REGION Network 31: Level Conveyors Tower 2 - SYSTEM 3
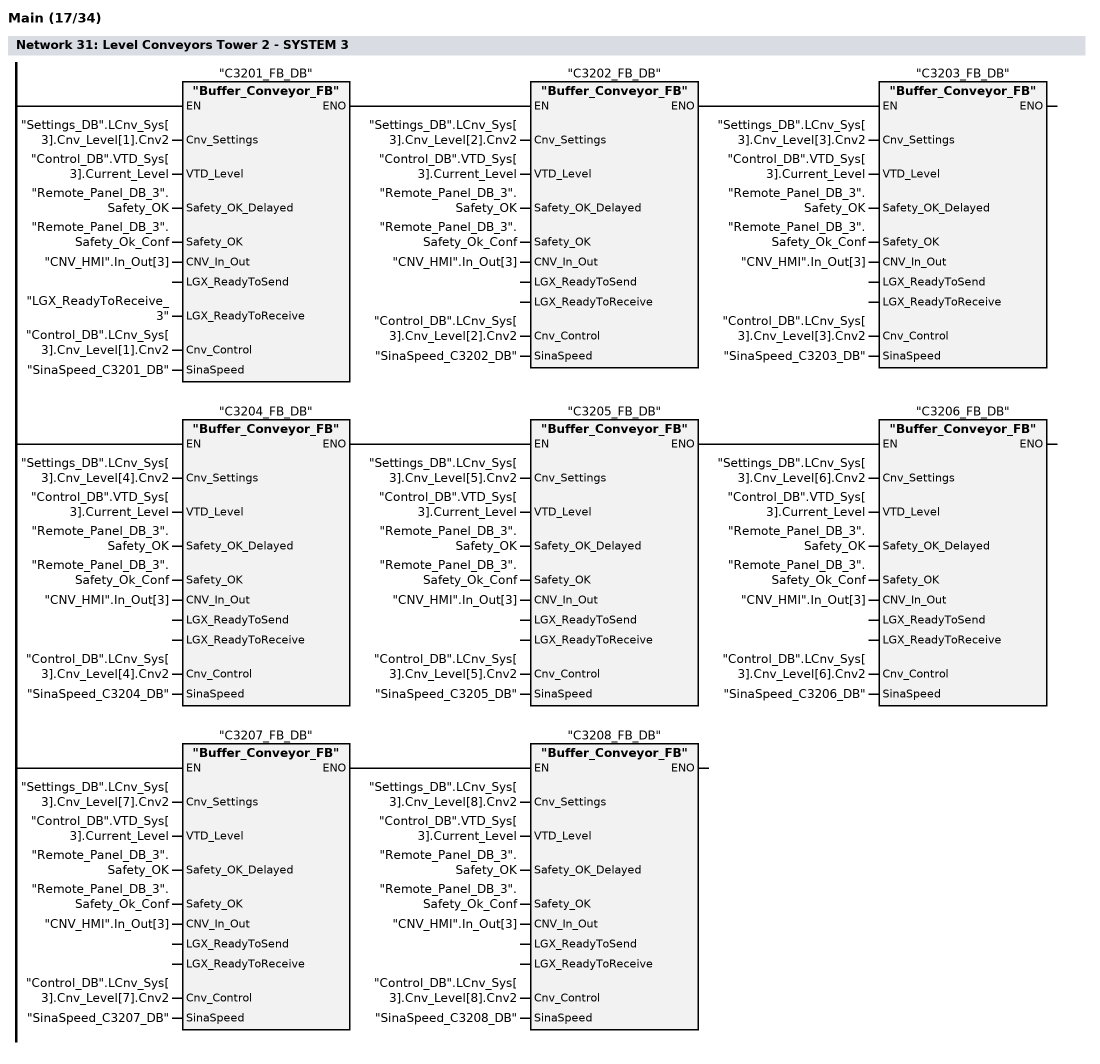
   RUNG wire#powerrail
      "C3201_FB_DB"(Cnv_Settings := "Settings_DB".LCnv_Sys[3].Cnv_Level[1].Cnv2, VTD_Level := "Control_DB".VTD_Sys[3].Current_Level, Safety_OK_Delayed := "Remote_Panel_DB_3".Safety_OK, Safety_OK := "Remote_Panel_DB_3".Safety_Ok_Conf, CNV_In_Out := "CNV_HMI".In_Out[3], LGX_ReadyToSend :=, LGX_ReadyToReceive := "LGX_ReadyToReceive_3", Cnv_Control := "Control_DB".LCnv_Sys[3].Cnv_Level[1].Cnv2, SinaSpeed := "SinaSpeed_C3201_DB")
      "C3202_FB_DB"(Cnv_Settings := "Settings_DB".LCnv_Sys[3].Cnv_Level[2].Cnv2, VTD_Level := "Control_DB".VTD_Sys[3].Current_Level, Safety_OK_Delayed := "Remote_Panel_DB_3".Safety_OK, Safety_OK := "Remote_Panel_DB_3".Safety_Ok_Conf, CNV_In_Out := "CNV_HMI".In_Out[3], LGX_ReadyToSend :=, LGX_ReadyToReceive :=, Cnv_Control := "Control_DB".LCnv_Sys[3].Cnv_Level[2].Cnv2, SinaSpeed := "SinaSpeed_C3202_DB")
      "C3203_FB_DB"(Cnv_Settings := "Settings_DB".LCnv_Sys[3].Cnv_Level[3].Cnv2, VTD_Level := "Control_DB".VTD_Sys[3].Current_Level, Safety_OK_Delayed := "Remote_Panel_DB_3".Safety_OK, Safety_OK := "Remote_Panel_DB_3".Safety_Ok_Conf, CNV_In_Out := "CNV_HMI".In_Out[3], LGX_ReadyToSend :=, LGX_ReadyToReceive :=, Cnv_Control := "Control_DB".LCnv_Sys[3].Cnv_Level[3].Cnv2, SinaSpeed := "SinaSpeed_C3203_DB")
   END_RUNG
   RUNG wire#powerrail
      "C3204_FB_DB"(Cnv_Settings := "Settings_DB".LCnv_Sys[3].Cnv_Level[4].Cnv2, VTD_Level := "Control_DB".VTD_Sys[3].Current_Level, Safety_OK_Delayed := "Remote_Panel_DB_3".Safety_OK, Safety_OK := "Remote_Panel_DB_3".Safety_Ok_Conf, CNV_In_Out := "CNV_HMI".In_Out[3], LGX_ReadyToSend :=, LGX_ReadyToReceive :=, Cnv_Control := "Control_DB".LCnv_Sys[3].Cnv_Level[4].Cnv2, SinaSpeed := "SinaSpeed_C3204_DB")
      "C3205_FB_DB"(Cnv_Settings := "Settings_DB".LCnv_Sys[3].Cnv_Level[5].Cnv2, VTD_Level := "Control_DB".VTD_Sys[3].Current_Level, Safety_OK_Delayed := "Remote_Panel_DB_3".Safety_OK, Safety_OK := "Remote_Panel_DB_3".Safety_Ok_Conf, CNV_In_Out := "CNV_HMI".In_Out[3], LGX_ReadyToSend :=, LGX_ReadyToReceive :=, Cnv_Control := "Control_DB".LCnv_Sys[3].Cnv_Level[5].Cnv2, SinaSpeed := "SinaSpeed_C3205_DB")
      "C3206_FB_DB"(Cnv_Settings := "Settings_DB".LCnv_Sys[3].Cnv_Level[6].Cnv2, VTD_Level := "Control_DB".VTD_Sys[3].Current_Level, Safety_OK_Delayed := "Remote_Panel_DB_3".Safety_OK, Safety_OK := "Remote_Panel_DB_3".Safety_Ok_Conf, CNV_In_Out := "CNV_HMI".In_Out[3], LGX_ReadyToSend :=, LGX_ReadyToReceive :=, Cnv_Control := "Control_DB".LCnv_Sys[3].Cnv_Level[6].Cnv2, SinaSpeed := "SinaSpeed_C3206_DB")
   END_RUNG
   RUNG wire#powerrail
      "C3207_FB_DB"(Cnv_Settings := "Settings_DB".LCnv_Sys[3].Cnv_Level[7].Cnv2, VTD_Level := "Control_DB".VTD_Sys[3].Current_Level, Safety_OK_Delayed := "Remote_Panel_DB_3".Safety_OK, Safety_OK := "Remote_Panel_DB_3".Safety_Ok_Conf, CNV_In_Out := "CNV_HMI".In_Out[3], LGX_ReadyToSend :=, LGX_ReadyToReceive :=, Cnv_Control := "Control_DB".LCnv_Sys[3].Cnv_Level[7].Cnv2, SinaSpeed := "SinaSpeed_C3207_DB")
      "C3208_FB_DB"(Cnv_Settings := "Settings_DB".LCnv_Sys[3].Cnv_Level[8].Cnv2, VTD_Level := "Control_DB".VTD_Sys[3].Current_Level, Safety_OK_Delayed := "Remote_Panel_DB_3".Safety_OK, Safety_OK := "Remote_Panel_DB_3".Safety_Ok_Conf, CNV_In_Out := "CNV_HMI".In_Out[3], LGX_ReadyToSend :=, LGX_ReadyToReceive :=, Cnv_Control := "Control_DB".LCnv_Sys[3].Cnv_Level[8].Cnv2, SinaSpeed := "SinaSpeed_C3208_DB")
   END_RUNG
   // the same network as SCL:
   "C3201_FB_DB"(Cnv_Settings := "Settings_DB".LCnv_Sys[3].Cnv_Level[1].Cnv2,   // "Buffer_Conveyor_FB"
                 VTD_Level := "Control_DB".VTD_Sys[3].Current_Level,
                 Safety_OK_Delayed := "Remote_Panel_DB_3".Safety_OK,
                 Safety_OK := "Remote_Panel_DB_3".Safety_Ok_Conf,
                 CNV_In_Out := "CNV_HMI".In_Out[3],
                 LGX_ReadyToReceive := "LGX_ReadyToReceive_3",
                 Cnv_Control := "Control_DB".LCnv_Sys[3].Cnv_Level[1].Cnv2,
                 SinaSpeed := "SinaSpeed_C3201_DB",
                 ENO => #_w1);
   "C3202_FB_DB"(EN := #_w1,   // "Buffer_Conveyor_FB"
                 Cnv_Settings := "Settings_DB".LCnv_Sys[3].Cnv_Level[2].Cnv2,
                 VTD_Level := "Control_DB".VTD_Sys[3].Current_Level,
                 Safety_OK_Delayed := "Remote_Panel_DB_3".Safety_OK,
                 Safety_OK := "Remote_Panel_DB_3".Safety_Ok_Conf,
                 CNV_In_Out := "CNV_HMI".In_Out[3],
                 Cnv_Control := "Control_DB".LCnv_Sys[3].Cnv_Level[2].Cnv2,
                 SinaSpeed := "SinaSpeed_C3202_DB",
                 ENO => #_w2);
   IF #_w2 THEN
       "C3203_FB_DB"(Cnv_Settings := "Settings_DB".LCnv_Sys[3].Cnv_Level[3].Cnv2,   // "Buffer_Conveyor_FB"
                     VTD_Level := "Control_DB".VTD_Sys[3].Current_Level,
                     Safety_OK_Delayed := "Remote_Panel_DB_3".Safety_OK,
                     Safety_OK := "Remote_Panel_DB_3".Safety_Ok_Conf,
                     CNV_In_Out := "CNV_HMI".In_Out[3],
                     Cnv_Control := "Control_DB".LCnv_Sys[3].Cnv_Level[3].Cnv2,
                     SinaSpeed := "SinaSpeed_C3203_DB");
   END_IF;
   "C3204_FB_DB"(Cnv_Settings := "Settings_DB".LCnv_Sys[3].Cnv_Level[4].Cnv2,   // "Buffer_Conveyor_FB"
                 VTD_Level := "Control_DB".VTD_Sys[3].Current_Level,
                 Safety_OK_Delayed := "Remote_Panel_DB_3".Safety_OK,
                 Safety_OK := "Remote_Panel_DB_3".Safety_Ok_Conf,
                 CNV_In_Out := "CNV_HMI".In_Out[3],
                 Cnv_Control := "Control_DB".LCnv_Sys[3].Cnv_Level[4].Cnv2,
                 SinaSpeed := "SinaSpeed_C3204_DB",
                 ENO => #_w3);
   "C3205_FB_DB"(EN := #_w3,   // "Buffer_Conveyor_FB"
                 Cnv_Settings := "Settings_DB".LCnv_Sys[3].Cnv_Level[5].Cnv2,
                 VTD_Level := "Control_DB".VTD_Sys[3].Current_Level,
                 Safety_OK_Delayed := "Remote_Panel_DB_3".Safety_OK,
                 Safety_OK := "Remote_Panel_DB_3".Safety_Ok_Conf,
                 CNV_In_Out := "CNV_HMI".In_Out[3],
                 Cnv_Control := "Control_DB".LCnv_Sys[3].Cnv_Level[5].Cnv2,
                 SinaSpeed := "SinaSpeed_C3205_DB",
                 ENO => #_w4);
   IF #_w4 THEN
       "C3206_FB_DB"(Cnv_Settings := "Settings_DB".LCnv_Sys[3].Cnv_Level[6].Cnv2,   // "Buffer_Conveyor_FB"
                     VTD_Level := "Control_DB".VTD_Sys[3].Current_Level,
                     Safety_OK_Delayed := "Remote_Panel_DB_3".Safety_OK,
                     Safety_OK := "Remote_Panel_DB_3".Safety_Ok_Conf,
                     CNV_In_Out := "CNV_HMI".In_Out[3],
                     Cnv_Control := "Control_DB".LCnv_Sys[3].Cnv_Level[6].Cnv2,
                     SinaSpeed := "SinaSpeed_C3206_DB");
   END_IF;
   "C3207_FB_DB"(Cnv_Settings := "Settings_DB".LCnv_Sys[3].Cnv_Level[7].Cnv2,   // "Buffer_Conveyor_FB"
                 VTD_Level := "Control_DB".VTD_Sys[3].Current_Level,
                 Safety_OK_Delayed := "Remote_Panel_DB_3".Safety_OK,
                 Safety_OK := "Remote_Panel_DB_3".Safety_Ok_Conf,
                 CNV_In_Out := "CNV_HMI".In_Out[3],
                 Cnv_Control := "Control_DB".LCnv_Sys[3].Cnv_Level[7].Cnv2,
                 SinaSpeed := "SinaSpeed_C3207_DB",
                 ENO => #_w5);
   IF #_w5 THEN
       "C3208_FB_DB"(Cnv_Settings := "Settings_DB".LCnv_Sys[3].Cnv_Level[8].Cnv2,   // "Buffer_Conveyor_FB"
                     VTD_Level := "Control_DB".VTD_Sys[3].Current_Level,
                     Safety_OK_Delayed := "Remote_Panel_DB_3".Safety_OK,
                     Safety_OK := "Remote_Panel_DB_3".Safety_Ok_Conf,
                     CNV_In_Out := "CNV_HMI".In_Out[3],
                     Cnv_Control := "Control_DB".LCnv_Sys[3].Cnv_Level[8].Cnv2,
                     SinaSpeed := "SinaSpeed_C3208_DB");
   END_IF;
END_REGION

REGION Network 32: SAFETY STOPPERS Tower 1 - SYSTEM 3
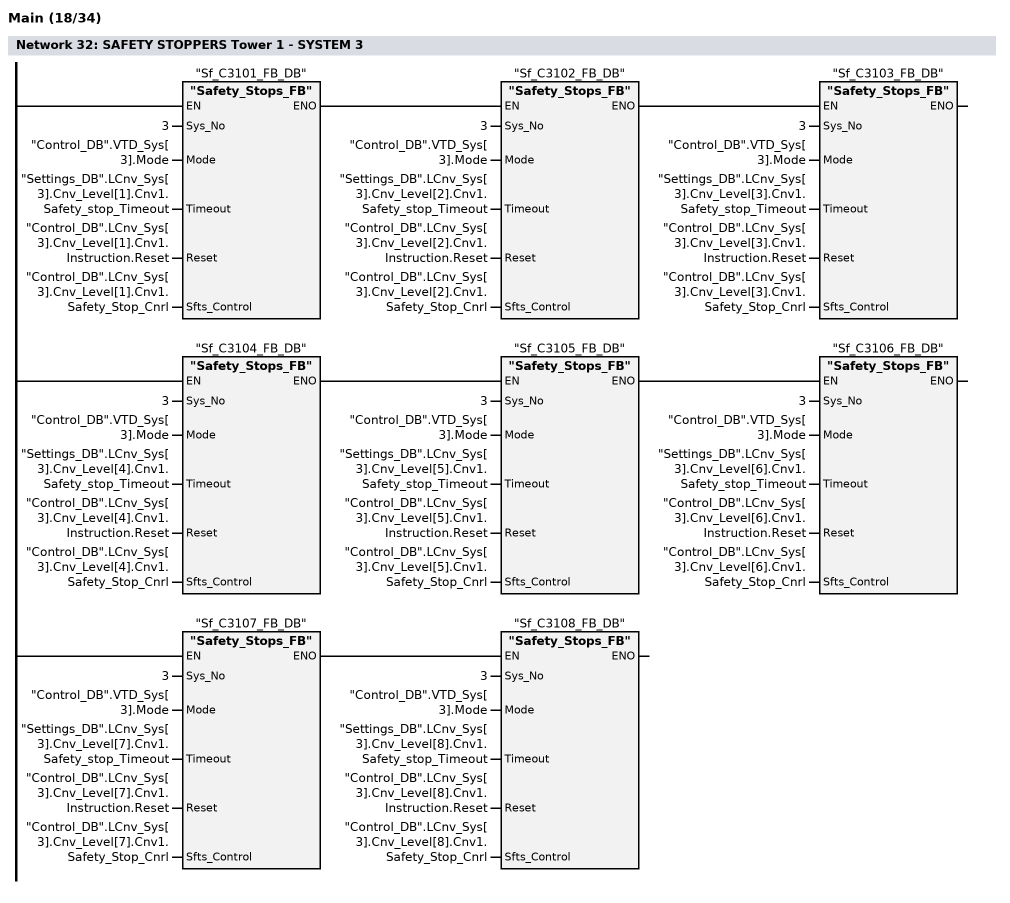
   RUNG wire#powerrail
      "Sf_C3101_FB_DB"(Sys_No := 3, Mode := "Control_DB".VTD_Sys[3].Mode, Timeout := "Settings_DB".LCnv_Sys[3].Cnv_Level[1].Cnv1.Safety_stop_Timeout, Reset := "Control_DB".LCnv_Sys[3].Cnv_Level[1].Cnv1.Instruction.Reset, Sfts_Control := "Control_DB".LCnv_Sys[3].Cnv_Level[1].Cnv1.Safety_Stop_Cnrl)
      "Sf_C3102_FB_DB"(Sys_No := 3, Mode := "Control_DB".VTD_Sys[3].Mode, Timeout := "Settings_DB".LCnv_Sys[3].Cnv_Level[2].Cnv1.Safety_stop_Timeout, Reset := "Control_DB".LCnv_Sys[3].Cnv_Level[2].Cnv1.Instruction.Reset, Sfts_Control := "Control_DB".LCnv_Sys[3].Cnv_Level[2].Cnv1.Safety_Stop_Cnrl)
      "Sf_C3103_FB_DB"(Sys_No := 3, Mode := "Control_DB".VTD_Sys[3].Mode, Timeout := "Settings_DB".LCnv_Sys[3].Cnv_Level[3].Cnv1.Safety_stop_Timeout, Reset := "Control_DB".LCnv_Sys[3].Cnv_Level[3].Cnv1.Instruction.Reset, Sfts_Control := "Control_DB".LCnv_Sys[3].Cnv_Level[3].Cnv1.Safety_Stop_Cnrl)
   END_RUNG
   RUNG wire#powerrail
      "Sf_C3104_FB_DB"(Sys_No := 3, Mode := "Control_DB".VTD_Sys[3].Mode, Timeout := "Settings_DB".LCnv_Sys[3].Cnv_Level[4].Cnv1.Safety_stop_Timeout, Reset := "Control_DB".LCnv_Sys[3].Cnv_Level[4].Cnv1.Instruction.Reset, Sfts_Control := "Control_DB".LCnv_Sys[3].Cnv_Level[4].Cnv1.Safety_Stop_Cnrl)
      "Sf_C3105_FB_DB"(Sys_No := 3, Mode := "Control_DB".VTD_Sys[3].Mode, Timeout := "Settings_DB".LCnv_Sys[3].Cnv_Level[5].Cnv1.Safety_stop_Timeout, Reset := "Control_DB".LCnv_Sys[3].Cnv_Level[5].Cnv1.Instruction.Reset, Sfts_Control := "Control_DB".LCnv_Sys[3].Cnv_Level[5].Cnv1.Safety_Stop_Cnrl)
      "Sf_C3106_FB_DB"(Sys_No := 3, Mode := "Control_DB".VTD_Sys[3].Mode, Timeout := "Settings_DB".LCnv_Sys[3].Cnv_Level[6].Cnv1.Safety_stop_Timeout, Reset := "Control_DB".LCnv_Sys[3].Cnv_Level[6].Cnv1.Instruction.Reset, Sfts_Control := "Control_DB".LCnv_Sys[3].Cnv_Level[6].Cnv1.Safety_Stop_Cnrl)
   END_RUNG
   RUNG wire#powerrail
      "Sf_C3107_FB_DB"(Sys_No := 3, Mode := "Control_DB".VTD_Sys[3].Mode, Timeout := "Settings_DB".LCnv_Sys[3].Cnv_Level[7].Cnv1.Safety_stop_Timeout, Reset := "Control_DB".LCnv_Sys[3].Cnv_Level[7].Cnv1.Instruction.Reset, Sfts_Control := "Control_DB".LCnv_Sys[3].Cnv_Level[7].Cnv1.Safety_Stop_Cnrl)
      "Sf_C3108_FB_DB"(Sys_No := 3, Mode := "Control_DB".VTD_Sys[3].Mode, Timeout := "Settings_DB".LCnv_Sys[3].Cnv_Level[8].Cnv1.Safety_stop_Timeout, Reset := "Control_DB".LCnv_Sys[3].Cnv_Level[8].Cnv1.Instruction.Reset, Sfts_Control := "Control_DB".LCnv_Sys[3].Cnv_Level[8].Cnv1.Safety_Stop_Cnrl)
   END_RUNG
   // the same network as SCL:
   "Sf_C3101_FB_DB"(Sys_No := 3,   // "Safety_Stops_FB"
                    Mode := "Control_DB".VTD_Sys[3].Mode,
                    Timeout := "Settings_DB".LCnv_Sys[3].Cnv_Level[1].Cnv1.Safety_stop_Timeout,
                    Reset := "Control_DB".LCnv_Sys[3].Cnv_Level[1].Cnv1.Instruction.Reset,
                    Sfts_Control := "Control_DB".LCnv_Sys[3].Cnv_Level[1].Cnv1.Safety_Stop_Cnrl,
                    ENO => #_w1);
   "Sf_C3102_FB_DB"(EN := #_w1,   // "Safety_Stops_FB"
                    Sys_No := 3,
                    Mode := "Control_DB".VTD_Sys[3].Mode,
                    Timeout := "Settings_DB".LCnv_Sys[3].Cnv_Level[2].Cnv1.Safety_stop_Timeout,
                    Reset := "Control_DB".LCnv_Sys[3].Cnv_Level[2].Cnv1.Instruction.Reset,
                    Sfts_Control := "Control_DB".LCnv_Sys[3].Cnv_Level[2].Cnv1.Safety_Stop_Cnrl,
                    ENO => #_w2);
   IF #_w2 THEN
       "Sf_C3103_FB_DB"(Sys_No := 3,   // "Safety_Stops_FB"
                        Mode := "Control_DB".VTD_Sys[3].Mode,
                        Timeout := "Settings_DB".LCnv_Sys[3].Cnv_Level[3].Cnv1.Safety_stop_Timeout,
                        Reset := "Control_DB".LCnv_Sys[3].Cnv_Level[3].Cnv1.Instruction.Reset,
                        Sfts_Control := "Control_DB".LCnv_Sys[3].Cnv_Level[3].Cnv1.Safety_Stop_Cnrl);
   END_IF;
   "Sf_C3104_FB_DB"(Sys_No := 3,   // "Safety_Stops_FB"
                    Mode := "Control_DB".VTD_Sys[3].Mode,
                    Timeout := "Settings_DB".LCnv_Sys[3].Cnv_Level[4].Cnv1.Safety_stop_Timeout,
                    Reset := "Control_DB".LCnv_Sys[3].Cnv_Level[4].Cnv1.Instruction.Reset,
                    Sfts_Control := "Control_DB".LCnv_Sys[3].Cnv_Level[4].Cnv1.Safety_Stop_Cnrl,
                    ENO => #_w3);
   "Sf_C3105_FB_DB"(EN := #_w3,   // "Safety_Stops_FB"
                    Sys_No := 3,
                    Mode := "Control_DB".VTD_Sys[3].Mode,
                    Timeout := "Settings_DB".LCnv_Sys[3].Cnv_Level[5].Cnv1.Safety_stop_Timeout,
                    Reset := "Control_DB".LCnv_Sys[3].Cnv_Level[5].Cnv1.Instruction.Reset,
                    Sfts_Control := "Control_DB".LCnv_Sys[3].Cnv_Level[5].Cnv1.Safety_Stop_Cnrl,
                    ENO => #_w4);
   IF #_w4 THEN
       "Sf_C3106_FB_DB"(Sys_No := 3,   // "Safety_Stops_FB"
                        Mode := "Control_DB".VTD_Sys[3].Mode,
                        Timeout := "Settings_DB".LCnv_Sys[3].Cnv_Level[6].Cnv1.Safety_stop_Timeout,
                        Reset := "Control_DB".LCnv_Sys[3].Cnv_Level[6].Cnv1.Instruction.Reset,
                        Sfts_Control := "Control_DB".LCnv_Sys[3].Cnv_Level[6].Cnv1.Safety_Stop_Cnrl);
   END_IF;
   "Sf_C3107_FB_DB"(Sys_No := 3,   // "Safety_Stops_FB"
                    Mode := "Control_DB".VTD_Sys[3].Mode,
                    Timeout := "Settings_DB".LCnv_Sys[3].Cnv_Level[7].Cnv1.Safety_stop_Timeout,
                    Reset := "Control_DB".LCnv_Sys[3].Cnv_Level[7].Cnv1.Instruction.Reset,
                    Sfts_Control := "Control_DB".LCnv_Sys[3].Cnv_Level[7].Cnv1.Safety_Stop_Cnrl,
                    ENO => #_w5);
   IF #_w5 THEN
       "Sf_C3108_FB_DB"(Sys_No := 3,   // "Safety_Stops_FB"
                        Mode := "Control_DB".VTD_Sys[3].Mode,
                        Timeout := "Settings_DB".LCnv_Sys[3].Cnv_Level[8].Cnv1.Safety_stop_Timeout,
                        Reset := "Control_DB".LCnv_Sys[3].Cnv_Level[8].Cnv1.Instruction.Reset,
                        Sfts_Control := "Control_DB".LCnv_Sys[3].Cnv_Level[8].Cnv1.Safety_Stop_Cnrl);
   END_IF;
END_REGION

REGION Network 33: SAFETY STOPPERS Tower 2 - SYSTEM 3
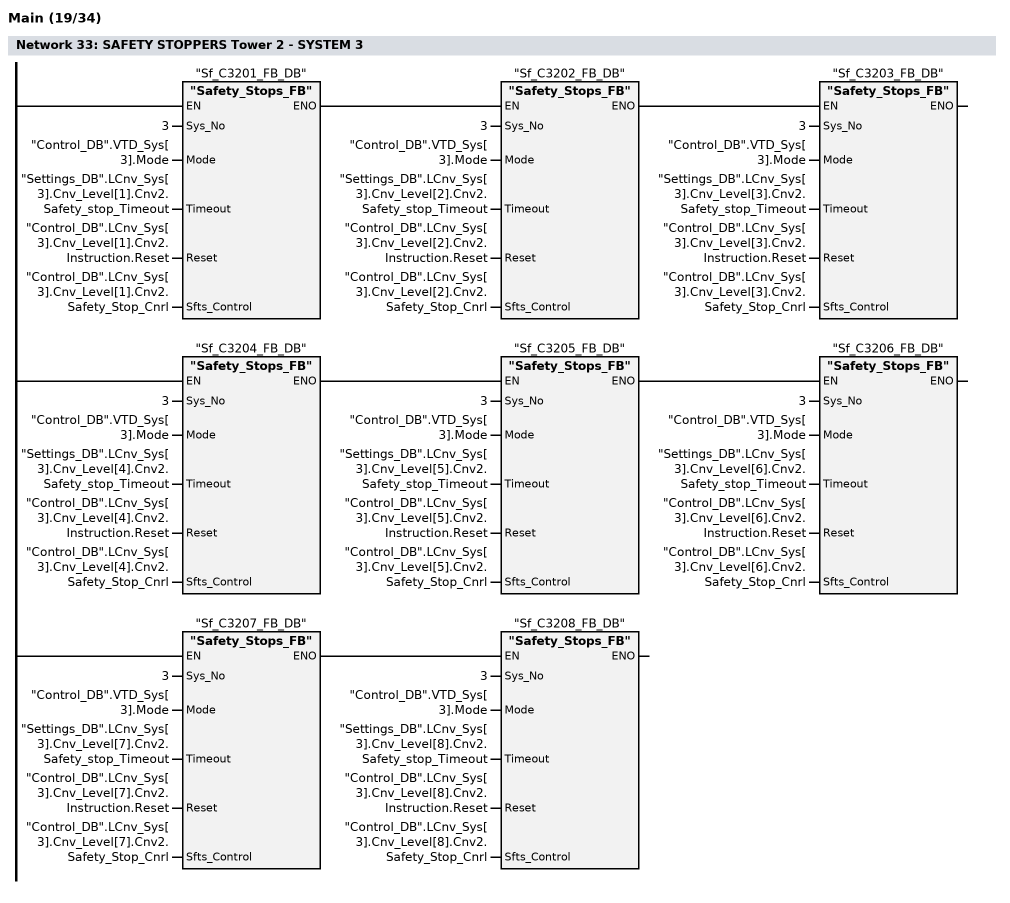
   RUNG wire#powerrail
      "Sf_C3201_FB_DB"(Sys_No := 3, Mode := "Control_DB".VTD_Sys[3].Mode, Timeout := "Settings_DB".LCnv_Sys[3].Cnv_Level[1].Cnv2.Safety_stop_Timeout, Reset := "Control_DB".LCnv_Sys[3].Cnv_Level[1].Cnv2.Instruction.Reset, Sfts_Control := "Control_DB".LCnv_Sys[3].Cnv_Level[1].Cnv2.Safety_Stop_Cnrl)
      "Sf_C3202_FB_DB"(Sys_No := 3, Mode := "Control_DB".VTD_Sys[3].Mode, Timeout := "Settings_DB".LCnv_Sys[3].Cnv_Level[2].Cnv2.Safety_stop_Timeout, Reset := "Control_DB".LCnv_Sys[3].Cnv_Level[2].Cnv2.Instruction.Reset, Sfts_Control := "Control_DB".LCnv_Sys[3].Cnv_Level[2].Cnv2.Safety_Stop_Cnrl)
      "Sf_C3203_FB_DB"(Sys_No := 3, Mode := "Control_DB".VTD_Sys[3].Mode, Timeout := "Settings_DB".LCnv_Sys[3].Cnv_Level[3].Cnv2.Safety_stop_Timeout, Reset := "Control_DB".LCnv_Sys[3].Cnv_Level[3].Cnv2.Instruction.Reset, Sfts_Control := "Control_DB".LCnv_Sys[3].Cnv_Level[3].Cnv2.Safety_Stop_Cnrl)
   END_RUNG
   RUNG wire#powerrail
      "Sf_C3204_FB_DB"(Sys_No := 3, Mode := "Control_DB".VTD_Sys[3].Mode, Timeout := "Settings_DB".LCnv_Sys[3].Cnv_Level[4].Cnv2.Safety_stop_Timeout, Reset := "Control_DB".LCnv_Sys[3].Cnv_Level[4].Cnv2.Instruction.Reset, Sfts_Control := "Control_DB".LCnv_Sys[3].Cnv_Level[4].Cnv2.Safety_Stop_Cnrl)
      "Sf_C3205_FB_DB"(Sys_No := 3, Mode := "Control_DB".VTD_Sys[3].Mode, Timeout := "Settings_DB".LCnv_Sys[3].Cnv_Level[5].Cnv2.Safety_stop_Timeout, Reset := "Control_DB".LCnv_Sys[3].Cnv_Level[5].Cnv2.Instruction.Reset, Sfts_Control := "Control_DB".LCnv_Sys[3].Cnv_Level[5].Cnv2.Safety_Stop_Cnrl)
      "Sf_C3206_FB_DB"(Sys_No := 3, Mode := "Control_DB".VTD_Sys[3].Mode, Timeout := "Settings_DB".LCnv_Sys[3].Cnv_Level[6].Cnv2.Safety_stop_Timeout, Reset := "Control_DB".LCnv_Sys[3].Cnv_Level[6].Cnv2.Instruction.Reset, Sfts_Control := "Control_DB".LCnv_Sys[3].Cnv_Level[6].Cnv2.Safety_Stop_Cnrl)
   END_RUNG
   RUNG wire#powerrail
      "Sf_C3207_FB_DB"(Sys_No := 3, Mode := "Control_DB".VTD_Sys[3].Mode, Timeout := "Settings_DB".LCnv_Sys[3].Cnv_Level[7].Cnv2.Safety_stop_Timeout, Reset := "Control_DB".LCnv_Sys[3].Cnv_Level[7].Cnv2.Instruction.Reset, Sfts_Control := "Control_DB".LCnv_Sys[3].Cnv_Level[7].Cnv2.Safety_Stop_Cnrl)
      "Sf_C3208_FB_DB"(Sys_No := 3, Mode := "Control_DB".VTD_Sys[3].Mode, Timeout := "Settings_DB".LCnv_Sys[3].Cnv_Level[8].Cnv2.Safety_stop_Timeout, Reset := "Control_DB".LCnv_Sys[3].Cnv_Level[8].Cnv2.Instruction.Reset, Sfts_Control := "Control_DB".LCnv_Sys[3].Cnv_Level[8].Cnv2.Safety_Stop_Cnrl)
   END_RUNG
   // the same network as SCL:
   "Sf_C3201_FB_DB"(Sys_No := 3,   // "Safety_Stops_FB"
                    Mode := "Control_DB".VTD_Sys[3].Mode,
                    Timeout := "Settings_DB".LCnv_Sys[3].Cnv_Level[1].Cnv2.Safety_stop_Timeout,
                    Reset := "Control_DB".LCnv_Sys[3].Cnv_Level[1].Cnv2.Instruction.Reset,
                    Sfts_Control := "Control_DB".LCnv_Sys[3].Cnv_Level[1].Cnv2.Safety_Stop_Cnrl,
                    ENO => #_w1);
   "Sf_C3202_FB_DB"(EN := #_w1,   // "Safety_Stops_FB"
                    Sys_No := 3,
                    Mode := "Control_DB".VTD_Sys[3].Mode,
                    Timeout := "Settings_DB".LCnv_Sys[3].Cnv_Level[2].Cnv2.Safety_stop_Timeout,
                    Reset := "Control_DB".LCnv_Sys[3].Cnv_Level[2].Cnv2.Instruction.Reset,
                    Sfts_Control := "Control_DB".LCnv_Sys[3].Cnv_Level[2].Cnv2.Safety_Stop_Cnrl,
                    ENO => #_w2);
   IF #_w2 THEN
       "Sf_C3203_FB_DB"(Sys_No := 3,   // "Safety_Stops_FB"
                        Mode := "Control_DB".VTD_Sys[3].Mode,
                        Timeout := "Settings_DB".LCnv_Sys[3].Cnv_Level[3].Cnv2.Safety_stop_Timeout,
                        Reset := "Control_DB".LCnv_Sys[3].Cnv_Level[3].Cnv2.Instruction.Reset,
                        Sfts_Control := "Control_DB".LCnv_Sys[3].Cnv_Level[3].Cnv2.Safety_Stop_Cnrl);
   END_IF;
   "Sf_C3204_FB_DB"(Sys_No := 3,   // "Safety_Stops_FB"
                    Mode := "Control_DB".VTD_Sys[3].Mode,
                    Timeout := "Settings_DB".LCnv_Sys[3].Cnv_Level[4].Cnv2.Safety_stop_Timeout,
                    Reset := "Control_DB".LCnv_Sys[3].Cnv_Level[4].Cnv2.Instruction.Reset,
                    Sfts_Control := "Control_DB".LCnv_Sys[3].Cnv_Level[4].Cnv2.Safety_Stop_Cnrl,
                    ENO => #_w3);
   "Sf_C3205_FB_DB"(EN := #_w3,   // "Safety_Stops_FB"
                    Sys_No := 3,
                    Mode := "Control_DB".VTD_Sys[3].Mode,
                    Timeout := "Settings_DB".LCnv_Sys[3].Cnv_Level[5].Cnv2.Safety_stop_Timeout,
                    Reset := "Control_DB".LCnv_Sys[3].Cnv_Level[5].Cnv2.Instruction.Reset,
                    Sfts_Control := "Control_DB".LCnv_Sys[3].Cnv_Level[5].Cnv2.Safety_Stop_Cnrl,
                    ENO => #_w4);
   IF #_w4 THEN
       "Sf_C3206_FB_DB"(Sys_No := 3,   // "Safety_Stops_FB"
                        Mode := "Control_DB".VTD_Sys[3].Mode,
                        Timeout := "Settings_DB".LCnv_Sys[3].Cnv_Level[6].Cnv2.Safety_stop_Timeout,
                        Reset := "Control_DB".LCnv_Sys[3].Cnv_Level[6].Cnv2.Instruction.Reset,
                        Sfts_Control := "Control_DB".LCnv_Sys[3].Cnv_Level[6].Cnv2.Safety_Stop_Cnrl);
   END_IF;
   "Sf_C3207_FB_DB"(Sys_No := 3,   // "Safety_Stops_FB"
                    Mode := "Control_DB".VTD_Sys[3].Mode,
                    Timeout := "Settings_DB".LCnv_Sys[3].Cnv_Level[7].Cnv2.Safety_stop_Timeout,
                    Reset := "Control_DB".LCnv_Sys[3].Cnv_Level[7].Cnv2.Instruction.Reset,
                    Sfts_Control := "Control_DB".LCnv_Sys[3].Cnv_Level[7].Cnv2.Safety_Stop_Cnrl,
                    ENO => #_w5);
   IF #_w5 THEN
       "Sf_C3208_FB_DB"(Sys_No := 3,   // "Safety_Stops_FB"
                        Mode := "Control_DB".VTD_Sys[3].Mode,
                        Timeout := "Settings_DB".LCnv_Sys[3].Cnv_Level[8].Cnv2.Safety_stop_Timeout,
                        Reset := "Control_DB".LCnv_Sys[3].Cnv_Level[8].Cnv2.Instruction.Reset,
                        Sfts_Control := "Control_DB".LCnv_Sys[3].Cnv_Level[8].Cnv2.Safety_Stop_Cnrl);
   END_IF;
END_REGION

REGION Network 34: SYSTEM 4
END_REGION

REGION Network 35: Level Conveyors Tower 1 - SYSTEM 4
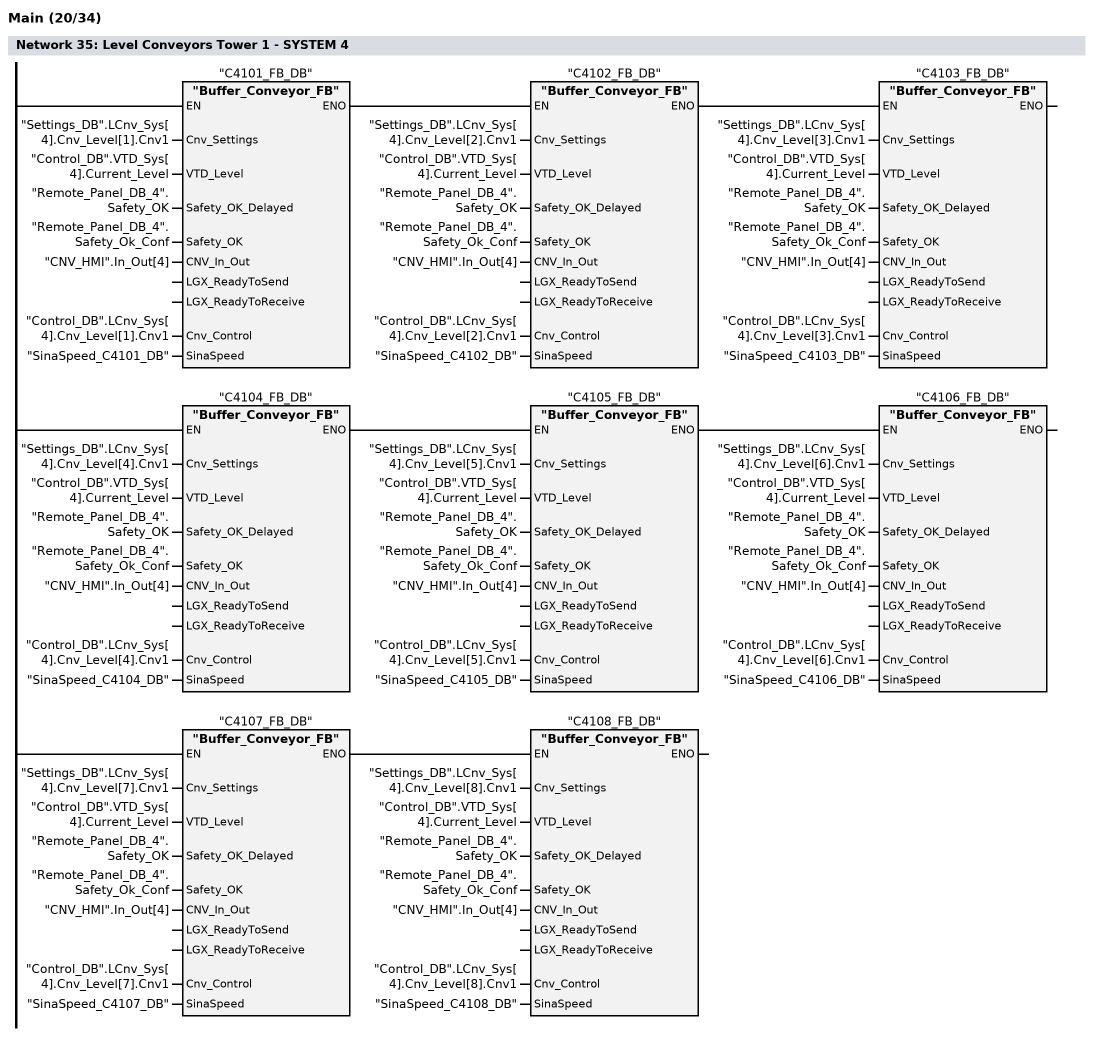
   RUNG wire#powerrail
      "C4101_FB_DB"(Cnv_Settings := "Settings_DB".LCnv_Sys[4].Cnv_Level[1].Cnv1, VTD_Level := "Control_DB".VTD_Sys[4].Current_Level, Safety_OK_Delayed := "Remote_Panel_DB_4".Safety_OK, Safety_OK := "Remote_Panel_DB_4".Safety_Ok_Conf, CNV_In_Out := "CNV_HMI".In_Out[4], LGX_ReadyToSend :=, LGX_ReadyToReceive :=, Cnv_Control := "Control_DB".LCnv_Sys[4].Cnv_Level[1].Cnv1, SinaSpeed := "SinaSpeed_C4101_DB")
      "C4102_FB_DB"(Cnv_Settings := "Settings_DB".LCnv_Sys[4].Cnv_Level[2].Cnv1, VTD_Level := "Control_DB".VTD_Sys[4].Current_Level, Safety_OK_Delayed := "Remote_Panel_DB_4".Safety_OK, Safety_OK := "Remote_Panel_DB_4".Safety_Ok_Conf, CNV_In_Out := "CNV_HMI".In_Out[4], LGX_ReadyToSend :=, LGX_ReadyToReceive :=, Cnv_Control := "Control_DB".LCnv_Sys[4].Cnv_Level[2].Cnv1, SinaSpeed := "SinaSpeed_C4102_DB")
      "C4103_FB_DB"(Cnv_Settings := "Settings_DB".LCnv_Sys[4].Cnv_Level[3].Cnv1, VTD_Level := "Control_DB".VTD_Sys[4].Current_Level, Safety_OK_Delayed := "Remote_Panel_DB_4".Safety_OK, Safety_OK := "Remote_Panel_DB_4".Safety_Ok_Conf, CNV_In_Out := "CNV_HMI".In_Out[4], LGX_ReadyToSend :=, LGX_ReadyToReceive :=, Cnv_Control := "Control_DB".LCnv_Sys[4].Cnv_Level[3].Cnv1, SinaSpeed := "SinaSpeed_C4103_DB")
   END_RUNG
   RUNG wire#powerrail
      "C4104_FB_DB"(Cnv_Settings := "Settings_DB".LCnv_Sys[4].Cnv_Level[4].Cnv1, VTD_Level := "Control_DB".VTD_Sys[4].Current_Level, Safety_OK_Delayed := "Remote_Panel_DB_4".Safety_OK, Safety_OK := "Remote_Panel_DB_4".Safety_Ok_Conf, CNV_In_Out := "CNV_HMI".In_Out[4], LGX_ReadyToSend :=, LGX_ReadyToReceive :=, Cnv_Control := "Control_DB".LCnv_Sys[4].Cnv_Level[4].Cnv1, SinaSpeed := "SinaSpeed_C4104_DB")
      "C4105_FB_DB"(Cnv_Settings := "Settings_DB".LCnv_Sys[4].Cnv_Level[5].Cnv1, VTD_Level := "Control_DB".VTD_Sys[4].Current_Level, Safety_OK_Delayed := "Remote_Panel_DB_4".Safety_OK, Safety_OK := "Remote_Panel_DB_4".Safety_Ok_Conf, CNV_In_Out := "CNV_HMI".In_Out[4], LGX_ReadyToSend :=, LGX_ReadyToReceive :=, Cnv_Control := "Control_DB".LCnv_Sys[4].Cnv_Level[5].Cnv1, SinaSpeed := "SinaSpeed_C4105_DB")
      "C4106_FB_DB"(Cnv_Settings := "Settings_DB".LCnv_Sys[4].Cnv_Level[6].Cnv1, VTD_Level := "Control_DB".VTD_Sys[4].Current_Level, Safety_OK_Delayed := "Remote_Panel_DB_4".Safety_OK, Safety_OK := "Remote_Panel_DB_4".Safety_Ok_Conf, CNV_In_Out := "CNV_HMI".In_Out[4], LGX_ReadyToSend :=, LGX_ReadyToReceive :=, Cnv_Control := "Control_DB".LCnv_Sys[4].Cnv_Level[6].Cnv1, SinaSpeed := "SinaSpeed_C4106_DB")
   END_RUNG
   RUNG wire#powerrail
      "C4107_FB_DB"(Cnv_Settings := "Settings_DB".LCnv_Sys[4].Cnv_Level[7].Cnv1, VTD_Level := "Control_DB".VTD_Sys[4].Current_Level, Safety_OK_Delayed := "Remote_Panel_DB_4".Safety_OK, Safety_OK := "Remote_Panel_DB_4".Safety_Ok_Conf, CNV_In_Out := "CNV_HMI".In_Out[4], LGX_ReadyToSend :=, LGX_ReadyToReceive :=, Cnv_Control := "Control_DB".LCnv_Sys[4].Cnv_Level[7].Cnv1, SinaSpeed := "SinaSpeed_C4107_DB")
      "C4108_FB_DB"(Cnv_Settings := "Settings_DB".LCnv_Sys[4].Cnv_Level[8].Cnv1, VTD_Level := "Control_DB".VTD_Sys[4].Current_Level, Safety_OK_Delayed := "Remote_Panel_DB_4".Safety_OK, Safety_OK := "Remote_Panel_DB_4".Safety_Ok_Conf, CNV_In_Out := "CNV_HMI".In_Out[4], LGX_ReadyToSend :=, LGX_ReadyToReceive :=, Cnv_Control := "Control_DB".LCnv_Sys[4].Cnv_Level[8].Cnv1, SinaSpeed := "SinaSpeed_C4108_DB")
   END_RUNG
   // the same network as SCL:
   "C4101_FB_DB"(Cnv_Settings := "Settings_DB".LCnv_Sys[4].Cnv_Level[1].Cnv1,   // "Buffer_Conveyor_FB"
                 VTD_Level := "Control_DB".VTD_Sys[4].Current_Level,
                 Safety_OK_Delayed := "Remote_Panel_DB_4".Safety_OK,
                 Safety_OK := "Remote_Panel_DB_4".Safety_Ok_Conf,
                 CNV_In_Out := "CNV_HMI".In_Out[4],
                 Cnv_Control := "Control_DB".LCnv_Sys[4].Cnv_Level[1].Cnv1,
                 SinaSpeed := "SinaSpeed_C4101_DB",
                 ENO => #_w1);
   "C4102_FB_DB"(EN := #_w1,   // "Buffer_Conveyor_FB"
                 Cnv_Settings := "Settings_DB".LCnv_Sys[4].Cnv_Level[2].Cnv1,
                 VTD_Level := "Control_DB".VTD_Sys[4].Current_Level,
                 Safety_OK_Delayed := "Remote_Panel_DB_4".Safety_OK,
                 Safety_OK := "Remote_Panel_DB_4".Safety_Ok_Conf,
                 CNV_In_Out := "CNV_HMI".In_Out[4],
                 Cnv_Control := "Control_DB".LCnv_Sys[4].Cnv_Level[2].Cnv1,
                 SinaSpeed := "SinaSpeed_C4102_DB",
                 ENO => #_w2);
   IF #_w2 THEN
       "C4103_FB_DB"(Cnv_Settings := "Settings_DB".LCnv_Sys[4].Cnv_Level[3].Cnv1,   // "Buffer_Conveyor_FB"
                     VTD_Level := "Control_DB".VTD_Sys[4].Current_Level,
                     Safety_OK_Delayed := "Remote_Panel_DB_4".Safety_OK,
                     Safety_OK := "Remote_Panel_DB_4".Safety_Ok_Conf,
                     CNV_In_Out := "CNV_HMI".In_Out[4],
                     Cnv_Control := "Control_DB".LCnv_Sys[4].Cnv_Level[3].Cnv1,
                     SinaSpeed := "SinaSpeed_C4103_DB");
   END_IF;
   "C4104_FB_DB"(Cnv_Settings := "Settings_DB".LCnv_Sys[4].Cnv_Level[4].Cnv1,   // "Buffer_Conveyor_FB"
                 VTD_Level := "Control_DB".VTD_Sys[4].Current_Level,
                 Safety_OK_Delayed := "Remote_Panel_DB_4".Safety_OK,
                 Safety_OK := "Remote_Panel_DB_4".Safety_Ok_Conf,
                 CNV_In_Out := "CNV_HMI".In_Out[4],
                 Cnv_Control := "Control_DB".LCnv_Sys[4].Cnv_Level[4].Cnv1,
                 SinaSpeed := "SinaSpeed_C4104_DB",
                 ENO => #_w3);
   "C4105_FB_DB"(EN := #_w3,   // "Buffer_Conveyor_FB"
                 Cnv_Settings := "Settings_DB".LCnv_Sys[4].Cnv_Level[5].Cnv1,
                 VTD_Level := "Control_DB".VTD_Sys[4].Current_Level,
                 Safety_OK_Delayed := "Remote_Panel_DB_4".Safety_OK,
                 Safety_OK := "Remote_Panel_DB_4".Safety_Ok_Conf,
                 CNV_In_Out := "CNV_HMI".In_Out[4],
                 Cnv_Control := "Control_DB".LCnv_Sys[4].Cnv_Level[5].Cnv1,
                 SinaSpeed := "SinaSpeed_C4105_DB",
                 ENO => #_w4);
   IF #_w4 THEN
       "C4106_FB_DB"(Cnv_Settings := "Settings_DB".LCnv_Sys[4].Cnv_Level[6].Cnv1,   // "Buffer_Conveyor_FB"
                     VTD_Level := "Control_DB".VTD_Sys[4].Current_Level,
                     Safety_OK_Delayed := "Remote_Panel_DB_4".Safety_OK,
                     Safety_OK := "Remote_Panel_DB_4".Safety_Ok_Conf,
                     CNV_In_Out := "CNV_HMI".In_Out[4],
                     Cnv_Control := "Control_DB".LCnv_Sys[4].Cnv_Level[6].Cnv1,
                     SinaSpeed := "SinaSpeed_C4106_DB");
   END_IF;
   "C4107_FB_DB"(Cnv_Settings := "Settings_DB".LCnv_Sys[4].Cnv_Level[7].Cnv1,   // "Buffer_Conveyor_FB"
                 VTD_Level := "Control_DB".VTD_Sys[4].Current_Level,
                 Safety_OK_Delayed := "Remote_Panel_DB_4".Safety_OK,
                 Safety_OK := "Remote_Panel_DB_4".Safety_Ok_Conf,
                 CNV_In_Out := "CNV_HMI".In_Out[4],
                 Cnv_Control := "Control_DB".LCnv_Sys[4].Cnv_Level[7].Cnv1,
                 SinaSpeed := "SinaSpeed_C4107_DB",
                 ENO => #_w5);
   IF #_w5 THEN
       "C4108_FB_DB"(Cnv_Settings := "Settings_DB".LCnv_Sys[4].Cnv_Level[8].Cnv1,   // "Buffer_Conveyor_FB"
                     VTD_Level := "Control_DB".VTD_Sys[4].Current_Level,
                     Safety_OK_Delayed := "Remote_Panel_DB_4".Safety_OK,
                     Safety_OK := "Remote_Panel_DB_4".Safety_Ok_Conf,
                     CNV_In_Out := "CNV_HMI".In_Out[4],
                     Cnv_Control := "Control_DB".LCnv_Sys[4].Cnv_Level[8].Cnv1,
                     SinaSpeed := "SinaSpeed_C4108_DB");
   END_IF;
END_REGION

REGION Network 36: SAFETY STOPPERS Tower 1 - SYSTEM 4
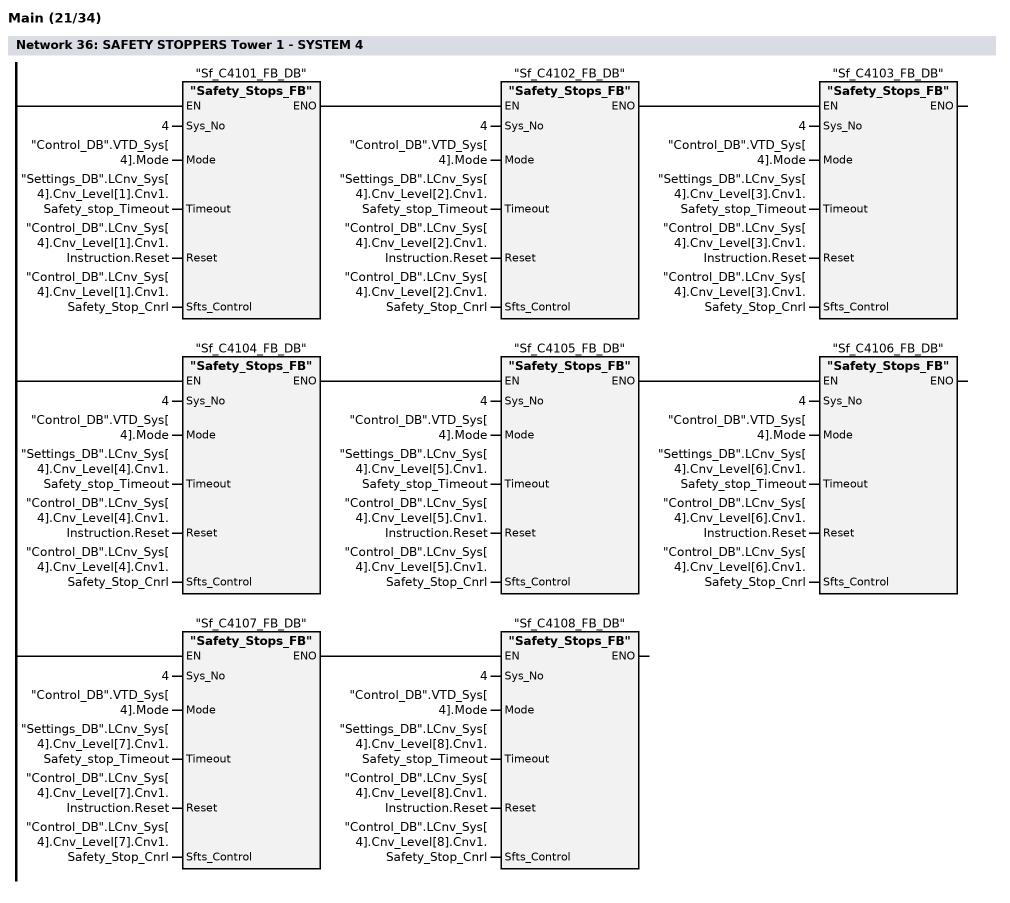
   RUNG wire#powerrail
      "Sf_C4101_FB_DB"(Sys_No := 4, Mode := "Control_DB".VTD_Sys[4].Mode, Timeout := "Settings_DB".LCnv_Sys[4].Cnv_Level[1].Cnv1.Safety_stop_Timeout, Reset := "Control_DB".LCnv_Sys[4].Cnv_Level[1].Cnv1.Instruction.Reset, Sfts_Control := "Control_DB".LCnv_Sys[4].Cnv_Level[1].Cnv1.Safety_Stop_Cnrl)
      "Sf_C4102_FB_DB"(Sys_No := 4, Mode := "Control_DB".VTD_Sys[4].Mode, Timeout := "Settings_DB".LCnv_Sys[4].Cnv_Level[2].Cnv1.Safety_stop_Timeout, Reset := "Control_DB".LCnv_Sys[4].Cnv_Level[2].Cnv1.Instruction.Reset, Sfts_Control := "Control_DB".LCnv_Sys[4].Cnv_Level[2].Cnv1.Safety_Stop_Cnrl)
      "Sf_C4103_FB_DB"(Sys_No := 4, Mode := "Control_DB".VTD_Sys[4].Mode, Timeout := "Settings_DB".LCnv_Sys[4].Cnv_Level[3].Cnv1.Safety_stop_Timeout, Reset := "Control_DB".LCnv_Sys[4].Cnv_Level[3].Cnv1.Instruction.Reset, Sfts_Control := "Control_DB".LCnv_Sys[4].Cnv_Level[3].Cnv1.Safety_Stop_Cnrl)
   END_RUNG
   RUNG wire#powerrail
      "Sf_C4104_FB_DB"(Sys_No := 4, Mode := "Control_DB".VTD_Sys[4].Mode, Timeout := "Settings_DB".LCnv_Sys[4].Cnv_Level[4].Cnv1.Safety_stop_Timeout, Reset := "Control_DB".LCnv_Sys[4].Cnv_Level[4].Cnv1.Instruction.Reset, Sfts_Control := "Control_DB".LCnv_Sys[4].Cnv_Level[4].Cnv1.Safety_Stop_Cnrl)
      "Sf_C4105_FB_DB"(Sys_No := 4, Mode := "Control_DB".VTD_Sys[4].Mode, Timeout := "Settings_DB".LCnv_Sys[4].Cnv_Level[5].Cnv1.Safety_stop_Timeout, Reset := "Control_DB".LCnv_Sys[4].Cnv_Level[5].Cnv1.Instruction.Reset, Sfts_Control := "Control_DB".LCnv_Sys[4].Cnv_Level[5].Cnv1.Safety_Stop_Cnrl)
      "Sf_C4106_FB_DB"(Sys_No := 4, Mode := "Control_DB".VTD_Sys[4].Mode, Timeout := "Settings_DB".LCnv_Sys[4].Cnv_Level[6].Cnv1.Safety_stop_Timeout, Reset := "Control_DB".LCnv_Sys[4].Cnv_Level[6].Cnv1.Instruction.Reset, Sfts_Control := "Control_DB".LCnv_Sys[4].Cnv_Level[6].Cnv1.Safety_Stop_Cnrl)
   END_RUNG
   RUNG wire#powerrail
      "Sf_C4107_FB_DB"(Sys_No := 4, Mode := "Control_DB".VTD_Sys[4].Mode, Timeout := "Settings_DB".LCnv_Sys[4].Cnv_Level[7].Cnv1.Safety_stop_Timeout, Reset := "Control_DB".LCnv_Sys[4].Cnv_Level[7].Cnv1.Instruction.Reset, Sfts_Control := "Control_DB".LCnv_Sys[4].Cnv_Level[7].Cnv1.Safety_Stop_Cnrl)
      "Sf_C4108_FB_DB"(Sys_No := 4, Mode := "Control_DB".VTD_Sys[4].Mode, Timeout := "Settings_DB".LCnv_Sys[4].Cnv_Level[8].Cnv1.Safety_stop_Timeout, Reset := "Control_DB".LCnv_Sys[4].Cnv_Level[8].Cnv1.Instruction.Reset, Sfts_Control := "Control_DB".LCnv_Sys[4].Cnv_Level[8].Cnv1.Safety_Stop_Cnrl)
   END_RUNG
   // the same network as SCL:
   "Sf_C4101_FB_DB"(Sys_No := 4,   // "Safety_Stops_FB"
                    Mode := "Control_DB".VTD_Sys[4].Mode,
                    Timeout := "Settings_DB".LCnv_Sys[4].Cnv_Level[1].Cnv1.Safety_stop_Timeout,
                    Reset := "Control_DB".LCnv_Sys[4].Cnv_Level[1].Cnv1.Instruction.Reset,
                    Sfts_Control := "Control_DB".LCnv_Sys[4].Cnv_Level[1].Cnv1.Safety_Stop_Cnrl,
                    ENO => #_w1);
   "Sf_C4102_FB_DB"(EN := #_w1,   // "Safety_Stops_FB"
                    Sys_No := 4,
                    Mode := "Control_DB".VTD_Sys[4].Mode,
                    Timeout := "Settings_DB".LCnv_Sys[4].Cnv_Level[2].Cnv1.Safety_stop_Timeout,
                    Reset := "Control_DB".LCnv_Sys[4].Cnv_Level[2].Cnv1.Instruction.Reset,
                    Sfts_Control := "Control_DB".LCnv_Sys[4].Cnv_Level[2].Cnv1.Safety_Stop_Cnrl,
                    ENO => #_w2);
   IF #_w2 THEN
       "Sf_C4103_FB_DB"(Sys_No := 4,   // "Safety_Stops_FB"
                        Mode := "Control_DB".VTD_Sys[4].Mode,
                        Timeout := "Settings_DB".LCnv_Sys[4].Cnv_Level[3].Cnv1.Safety_stop_Timeout,
                        Reset := "Control_DB".LCnv_Sys[4].Cnv_Level[3].Cnv1.Instruction.Reset,
                        Sfts_Control := "Control_DB".LCnv_Sys[4].Cnv_Level[3].Cnv1.Safety_Stop_Cnrl);
   END_IF;
   "Sf_C4104_FB_DB"(Sys_No := 4,   // "Safety_Stops_FB"
                    Mode := "Control_DB".VTD_Sys[4].Mode,
                    Timeout := "Settings_DB".LCnv_Sys[4].Cnv_Level[4].Cnv1.Safety_stop_Timeout,
                    Reset := "Control_DB".LCnv_Sys[4].Cnv_Level[4].Cnv1.Instruction.Reset,
                    Sfts_Control := "Control_DB".LCnv_Sys[4].Cnv_Level[4].Cnv1.Safety_Stop_Cnrl,
                    ENO => #_w3);
   "Sf_C4105_FB_DB"(EN := #_w3,   // "Safety_Stops_FB"
                    Sys_No := 4,
                    Mode := "Control_DB".VTD_Sys[4].Mode,
                    Timeout := "Settings_DB".LCnv_Sys[4].Cnv_Level[5].Cnv1.Safety_stop_Timeout,
                    Reset := "Control_DB".LCnv_Sys[4].Cnv_Level[5].Cnv1.Instruction.Reset,
                    Sfts_Control := "Control_DB".LCnv_Sys[4].Cnv_Level[5].Cnv1.Safety_Stop_Cnrl,
                    ENO => #_w4);
   IF #_w4 THEN
       "Sf_C4106_FB_DB"(Sys_No := 4,   // "Safety_Stops_FB"
                        Mode := "Control_DB".VTD_Sys[4].Mode,
                        Timeout := "Settings_DB".LCnv_Sys[4].Cnv_Level[6].Cnv1.Safety_stop_Timeout,
                        Reset := "Control_DB".LCnv_Sys[4].Cnv_Level[6].Cnv1.Instruction.Reset,
                        Sfts_Control := "Control_DB".LCnv_Sys[4].Cnv_Level[6].Cnv1.Safety_Stop_Cnrl);
   END_IF;
   "Sf_C4107_FB_DB"(Sys_No := 4,   // "Safety_Stops_FB"
                    Mode := "Control_DB".VTD_Sys[4].Mode,
                    Timeout := "Settings_DB".LCnv_Sys[4].Cnv_Level[7].Cnv1.Safety_stop_Timeout,
                    Reset := "Control_DB".LCnv_Sys[4].Cnv_Level[7].Cnv1.Instruction.Reset,
                    Sfts_Control := "Control_DB".LCnv_Sys[4].Cnv_Level[7].Cnv1.Safety_Stop_Cnrl,
                    ENO => #_w5);
   IF #_w5 THEN
       "Sf_C4108_FB_DB"(Sys_No := 4,   // "Safety_Stops_FB"
                        Mode := "Control_DB".VTD_Sys[4].Mode,
                        Timeout := "Settings_DB".LCnv_Sys[4].Cnv_Level[8].Cnv1.Safety_stop_Timeout,
                        Reset := "Control_DB".LCnv_Sys[4].Cnv_Level[8].Cnv1.Instruction.Reset,
                        Sfts_Control := "Control_DB".LCnv_Sys[4].Cnv_Level[8].Cnv1.Safety_Stop_Cnrl);
   END_IF;
END_REGION

REGION Network 37: SYSTEM 5
END_REGION

REGION Network 38: Level Conveyors Tower 1 - SYSTEM 5
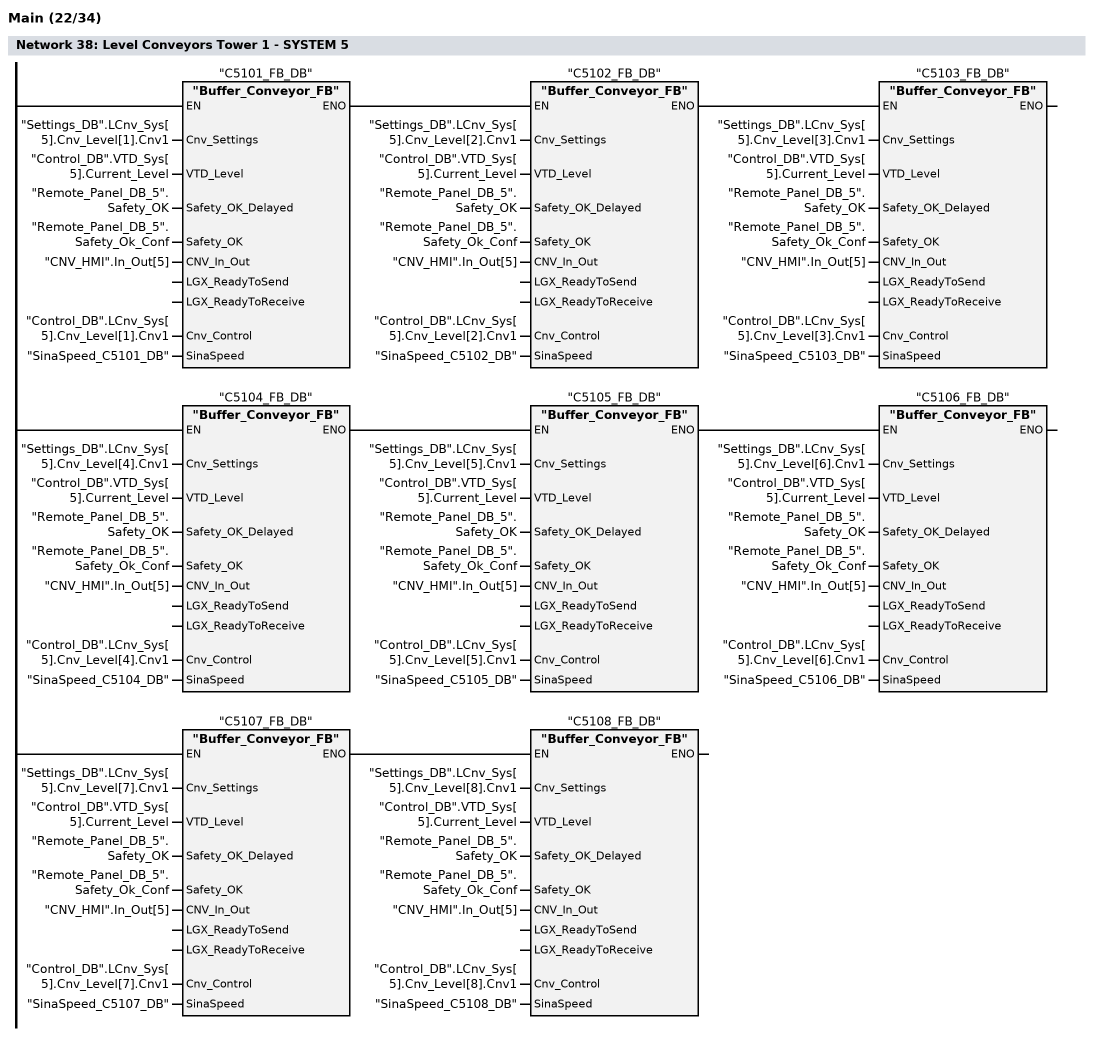
   RUNG wire#powerrail
      "C5101_FB_DB"(Cnv_Settings := "Settings_DB".LCnv_Sys[5].Cnv_Level[1].Cnv1, VTD_Level := "Control_DB".VTD_Sys[5].Current_Level, Safety_OK_Delayed := "Remote_Panel_DB_5".Safety_OK, Safety_OK := "Remote_Panel_DB_5".Safety_Ok_Conf, CNV_In_Out := "CNV_HMI".In_Out[5], LGX_ReadyToSend :=, LGX_ReadyToReceive :=, Cnv_Control := "Control_DB".LCnv_Sys[5].Cnv_Level[1].Cnv1, SinaSpeed := "SinaSpeed_C5101_DB")
      "C5102_FB_DB"(Cnv_Settings := "Settings_DB".LCnv_Sys[5].Cnv_Level[2].Cnv1, VTD_Level := "Control_DB".VTD_Sys[5].Current_Level, Safety_OK_Delayed := "Remote_Panel_DB_5".Safety_OK, Safety_OK := "Remote_Panel_DB_5".Safety_Ok_Conf, CNV_In_Out := "CNV_HMI".In_Out[5], LGX_ReadyToSend :=, LGX_ReadyToReceive :=, Cnv_Control := "Control_DB".LCnv_Sys[5].Cnv_Level[2].Cnv1, SinaSpeed := "SinaSpeed_C5102_DB")
      "C5103_FB_DB"(Cnv_Settings := "Settings_DB".LCnv_Sys[5].Cnv_Level[3].Cnv1, VTD_Level := "Control_DB".VTD_Sys[5].Current_Level, Safety_OK_Delayed := "Remote_Panel_DB_5".Safety_OK, Safety_OK := "Remote_Panel_DB_5".Safety_Ok_Conf, CNV_In_Out := "CNV_HMI".In_Out[5], LGX_ReadyToSend :=, LGX_ReadyToReceive :=, Cnv_Control := "Control_DB".LCnv_Sys[5].Cnv_Level[3].Cnv1, SinaSpeed := "SinaSpeed_C5103_DB")
   END_RUNG
   RUNG wire#powerrail
      "C5104_FB_DB"(Cnv_Settings := "Settings_DB".LCnv_Sys[5].Cnv_Level[4].Cnv1, VTD_Level := "Control_DB".VTD_Sys[5].Current_Level, Safety_OK_Delayed := "Remote_Panel_DB_5".Safety_OK, Safety_OK := "Remote_Panel_DB_5".Safety_Ok_Conf, CNV_In_Out := "CNV_HMI".In_Out[5], LGX_ReadyToSend :=, LGX_ReadyToReceive :=, Cnv_Control := "Control_DB".LCnv_Sys[5].Cnv_Level[4].Cnv1, SinaSpeed := "SinaSpeed_C5104_DB")
      "C5105_FB_DB"(Cnv_Settings := "Settings_DB".LCnv_Sys[5].Cnv_Level[5].Cnv1, VTD_Level := "Control_DB".VTD_Sys[5].Current_Level, Safety_OK_Delayed := "Remote_Panel_DB_5".Safety_OK, Safety_OK := "Remote_Panel_DB_5".Safety_Ok_Conf, CNV_In_Out := "CNV_HMI".In_Out[5], LGX_ReadyToSend :=, LGX_ReadyToReceive :=, Cnv_Control := "Control_DB".LCnv_Sys[5].Cnv_Level[5].Cnv1, SinaSpeed := "SinaSpeed_C5105_DB")
      "C5106_FB_DB"(Cnv_Settings := "Settings_DB".LCnv_Sys[5].Cnv_Level[6].Cnv1, VTD_Level := "Control_DB".VTD_Sys[5].Current_Level, Safety_OK_Delayed := "Remote_Panel_DB_5".Safety_OK, Safety_OK := "Remote_Panel_DB_5".Safety_Ok_Conf, CNV_In_Out := "CNV_HMI".In_Out[5], LGX_ReadyToSend :=, LGX_ReadyToReceive :=, Cnv_Control := "Control_DB".LCnv_Sys[5].Cnv_Level[6].Cnv1, SinaSpeed := "SinaSpeed_C5106_DB")
   END_RUNG
   RUNG wire#powerrail
      "C5107_FB_DB"(Cnv_Settings := "Settings_DB".LCnv_Sys[5].Cnv_Level[7].Cnv1, VTD_Level := "Control_DB".VTD_Sys[5].Current_Level, Safety_OK_Delayed := "Remote_Panel_DB_5".Safety_OK, Safety_OK := "Remote_Panel_DB_5".Safety_Ok_Conf, CNV_In_Out := "CNV_HMI".In_Out[5], LGX_ReadyToSend :=, LGX_ReadyToReceive :=, Cnv_Control := "Control_DB".LCnv_Sys[5].Cnv_Level[7].Cnv1, SinaSpeed := "SinaSpeed_C5107_DB")
      "C5108_FB_DB"(Cnv_Settings := "Settings_DB".LCnv_Sys[5].Cnv_Level[8].Cnv1, VTD_Level := "Control_DB".VTD_Sys[5].Current_Level, Safety_OK_Delayed := "Remote_Panel_DB_5".Safety_OK, Safety_OK := "Remote_Panel_DB_5".Safety_Ok_Conf, CNV_In_Out := "CNV_HMI".In_Out[5], LGX_ReadyToSend :=, LGX_ReadyToReceive :=, Cnv_Control := "Control_DB".LCnv_Sys[5].Cnv_Level[8].Cnv1, SinaSpeed := "SinaSpeed_C5108_DB")
   END_RUNG
   // the same network as SCL:
   "C5101_FB_DB"(Cnv_Settings := "Settings_DB".LCnv_Sys[5].Cnv_Level[1].Cnv1,   // "Buffer_Conveyor_FB"
                 VTD_Level := "Control_DB".VTD_Sys[5].Current_Level,
                 Safety_OK_Delayed := "Remote_Panel_DB_5".Safety_OK,
                 Safety_OK := "Remote_Panel_DB_5".Safety_Ok_Conf,
                 CNV_In_Out := "CNV_HMI".In_Out[5],
                 Cnv_Control := "Control_DB".LCnv_Sys[5].Cnv_Level[1].Cnv1,
                 SinaSpeed := "SinaSpeed_C5101_DB",
                 ENO => #_w1);
   "C5102_FB_DB"(EN := #_w1,   // "Buffer_Conveyor_FB"
                 Cnv_Settings := "Settings_DB".LCnv_Sys[5].Cnv_Level[2].Cnv1,
                 VTD_Level := "Control_DB".VTD_Sys[5].Current_Level,
                 Safety_OK_Delayed := "Remote_Panel_DB_5".Safety_OK,
                 Safety_OK := "Remote_Panel_DB_5".Safety_Ok_Conf,
                 CNV_In_Out := "CNV_HMI".In_Out[5],
                 Cnv_Control := "Control_DB".LCnv_Sys[5].Cnv_Level[2].Cnv1,
                 SinaSpeed := "SinaSpeed_C5102_DB",
                 ENO => #_w2);
   IF #_w2 THEN
       "C5103_FB_DB"(Cnv_Settings := "Settings_DB".LCnv_Sys[5].Cnv_Level[3].Cnv1,   // "Buffer_Conveyor_FB"
                     VTD_Level := "Control_DB".VTD_Sys[5].Current_Level,
                     Safety_OK_Delayed := "Remote_Panel_DB_5".Safety_OK,
                     Safety_OK := "Remote_Panel_DB_5".Safety_Ok_Conf,
                     CNV_In_Out := "CNV_HMI".In_Out[5],
                     Cnv_Control := "Control_DB".LCnv_Sys[5].Cnv_Level[3].Cnv1,
                     SinaSpeed := "SinaSpeed_C5103_DB");
   END_IF;
   "C5104_FB_DB"(Cnv_Settings := "Settings_DB".LCnv_Sys[5].Cnv_Level[4].Cnv1,   // "Buffer_Conveyor_FB"
                 VTD_Level := "Control_DB".VTD_Sys[5].Current_Level,
                 Safety_OK_Delayed := "Remote_Panel_DB_5".Safety_OK,
                 Safety_OK := "Remote_Panel_DB_5".Safety_Ok_Conf,
                 CNV_In_Out := "CNV_HMI".In_Out[5],
                 Cnv_Control := "Control_DB".LCnv_Sys[5].Cnv_Level[4].Cnv1,
                 SinaSpeed := "SinaSpeed_C5104_DB",
                 ENO => #_w3);
   "C5105_FB_DB"(EN := #_w3,   // "Buffer_Conveyor_FB"
                 Cnv_Settings := "Settings_DB".LCnv_Sys[5].Cnv_Level[5].Cnv1,
                 VTD_Level := "Control_DB".VTD_Sys[5].Current_Level,
                 Safety_OK_Delayed := "Remote_Panel_DB_5".Safety_OK,
                 Safety_OK := "Remote_Panel_DB_5".Safety_Ok_Conf,
                 CNV_In_Out := "CNV_HMI".In_Out[5],
                 Cnv_Control := "Control_DB".LCnv_Sys[5].Cnv_Level[5].Cnv1,
                 SinaSpeed := "SinaSpeed_C5105_DB",
                 ENO => #_w4);
   IF #_w4 THEN
       "C5106_FB_DB"(Cnv_Settings := "Settings_DB".LCnv_Sys[5].Cnv_Level[6].Cnv1,   // "Buffer_Conveyor_FB"
                     VTD_Level := "Control_DB".VTD_Sys[5].Current_Level,
                     Safety_OK_Delayed := "Remote_Panel_DB_5".Safety_OK,
                     Safety_OK := "Remote_Panel_DB_5".Safety_Ok_Conf,
                     CNV_In_Out := "CNV_HMI".In_Out[5],
                     Cnv_Control := "Control_DB".LCnv_Sys[5].Cnv_Level[6].Cnv1,
                     SinaSpeed := "SinaSpeed_C5106_DB");
   END_IF;
   "C5107_FB_DB"(Cnv_Settings := "Settings_DB".LCnv_Sys[5].Cnv_Level[7].Cnv1,   // "Buffer_Conveyor_FB"
                 VTD_Level := "Control_DB".VTD_Sys[5].Current_Level,
                 Safety_OK_Delayed := "Remote_Panel_DB_5".Safety_OK,
                 Safety_OK := "Remote_Panel_DB_5".Safety_Ok_Conf,
                 CNV_In_Out := "CNV_HMI".In_Out[5],
                 Cnv_Control := "Control_DB".LCnv_Sys[5].Cnv_Level[7].Cnv1,
                 SinaSpeed := "SinaSpeed_C5107_DB",
                 ENO => #_w5);
   IF #_w5 THEN
       "C5108_FB_DB"(Cnv_Settings := "Settings_DB".LCnv_Sys[5].Cnv_Level[8].Cnv1,   // "Buffer_Conveyor_FB"
                     VTD_Level := "Control_DB".VTD_Sys[5].Current_Level,
                     Safety_OK_Delayed := "Remote_Panel_DB_5".Safety_OK,
                     Safety_OK := "Remote_Panel_DB_5".Safety_Ok_Conf,
                     CNV_In_Out := "CNV_HMI".In_Out[5],
                     Cnv_Control := "Control_DB".LCnv_Sys[5].Cnv_Level[8].Cnv1,
                     SinaSpeed := "SinaSpeed_C5108_DB");
   END_IF;
END_REGION

REGION Network 39: SAFETY STOPPERS Tower 1 - SYSTEM 5
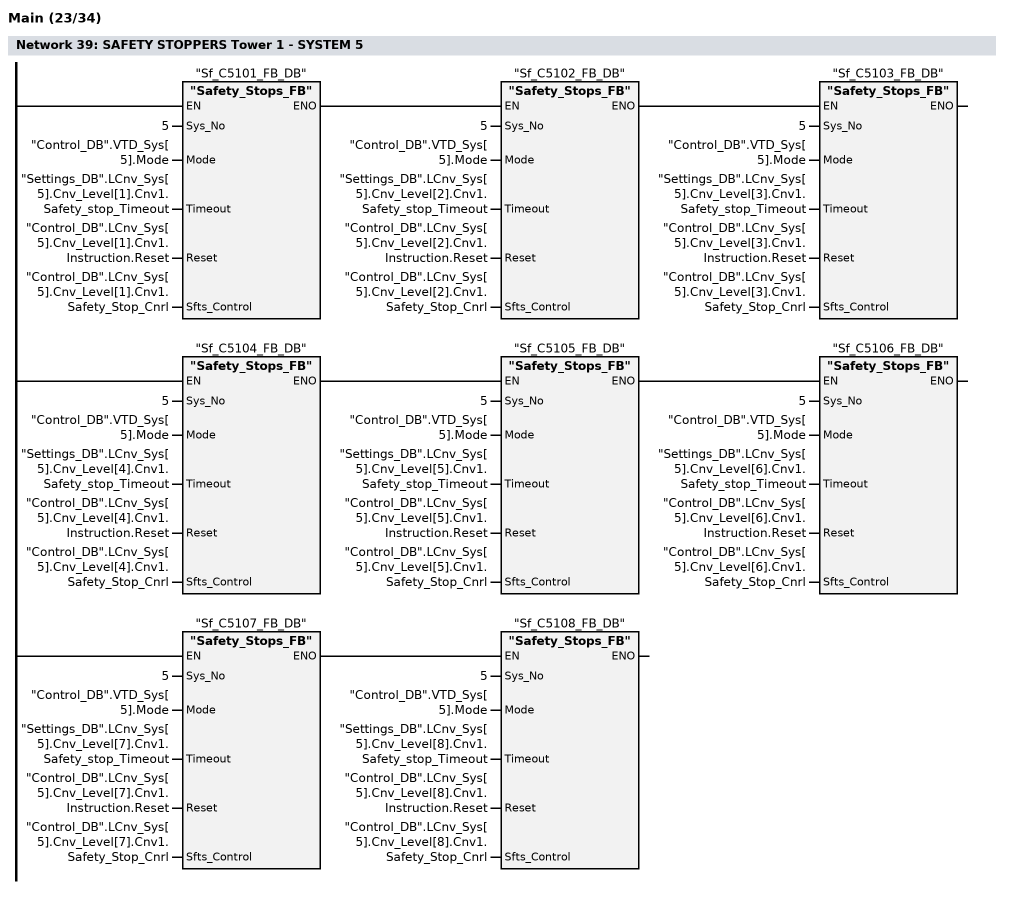
   RUNG wire#powerrail
      "Sf_C5101_FB_DB"(Sys_No := 5, Mode := "Control_DB".VTD_Sys[5].Mode, Timeout := "Settings_DB".LCnv_Sys[5].Cnv_Level[1].Cnv1.Safety_stop_Timeout, Reset := "Control_DB".LCnv_Sys[5].Cnv_Level[1].Cnv1.Instruction.Reset, Sfts_Control := "Control_DB".LCnv_Sys[5].Cnv_Level[1].Cnv1.Safety_Stop_Cnrl)
      "Sf_C5102_FB_DB"(Sys_No := 5, Mode := "Control_DB".VTD_Sys[5].Mode, Timeout := "Settings_DB".LCnv_Sys[5].Cnv_Level[2].Cnv1.Safety_stop_Timeout, Reset := "Control_DB".LCnv_Sys[5].Cnv_Level[2].Cnv1.Instruction.Reset, Sfts_Control := "Control_DB".LCnv_Sys[5].Cnv_Level[2].Cnv1.Safety_Stop_Cnrl)
      "Sf_C5103_FB_DB"(Sys_No := 5, Mode := "Control_DB".VTD_Sys[5].Mode, Timeout := "Settings_DB".LCnv_Sys[5].Cnv_Level[3].Cnv1.Safety_stop_Timeout, Reset := "Control_DB".LCnv_Sys[5].Cnv_Level[3].Cnv1.Instruction.Reset, Sfts_Control := "Control_DB".LCnv_Sys[5].Cnv_Level[3].Cnv1.Safety_Stop_Cnrl)
   END_RUNG
   RUNG wire#powerrail
      "Sf_C5104_FB_DB"(Sys_No := 5, Mode := "Control_DB".VTD_Sys[5].Mode, Timeout := "Settings_DB".LCnv_Sys[5].Cnv_Level[4].Cnv1.Safety_stop_Timeout, Reset := "Control_DB".LCnv_Sys[5].Cnv_Level[4].Cnv1.Instruction.Reset, Sfts_Control := "Control_DB".LCnv_Sys[5].Cnv_Level[4].Cnv1.Safety_Stop_Cnrl)
      "Sf_C5105_FB_DB"(Sys_No := 5, Mode := "Control_DB".VTD_Sys[5].Mode, Timeout := "Settings_DB".LCnv_Sys[5].Cnv_Level[5].Cnv1.Safety_stop_Timeout, Reset := "Control_DB".LCnv_Sys[5].Cnv_Level[5].Cnv1.Instruction.Reset, Sfts_Control := "Control_DB".LCnv_Sys[5].Cnv_Level[5].Cnv1.Safety_Stop_Cnrl)
      "Sf_C5106_FB_DB"(Sys_No := 5, Mode := "Control_DB".VTD_Sys[5].Mode, Timeout := "Settings_DB".LCnv_Sys[5].Cnv_Level[6].Cnv1.Safety_stop_Timeout, Reset := "Control_DB".LCnv_Sys[5].Cnv_Level[6].Cnv1.Instruction.Reset, Sfts_Control := "Control_DB".LCnv_Sys[5].Cnv_Level[6].Cnv1.Safety_Stop_Cnrl)
   END_RUNG
   RUNG wire#powerrail
      "Sf_C5107_FB_DB"(Sys_No := 5, Mode := "Control_DB".VTD_Sys[5].Mode, Timeout := "Settings_DB".LCnv_Sys[5].Cnv_Level[7].Cnv1.Safety_stop_Timeout, Reset := "Control_DB".LCnv_Sys[5].Cnv_Level[7].Cnv1.Instruction.Reset, Sfts_Control := "Control_DB".LCnv_Sys[5].Cnv_Level[7].Cnv1.Safety_Stop_Cnrl)
      "Sf_C5108_FB_DB"(Sys_No := 5, Mode := "Control_DB".VTD_Sys[5].Mode, Timeout := "Settings_DB".LCnv_Sys[5].Cnv_Level[8].Cnv1.Safety_stop_Timeout, Reset := "Control_DB".LCnv_Sys[5].Cnv_Level[8].Cnv1.Instruction.Reset, Sfts_Control := "Control_DB".LCnv_Sys[5].Cnv_Level[8].Cnv1.Safety_Stop_Cnrl)
   END_RUNG
   // the same network as SCL:
   "Sf_C5101_FB_DB"(Sys_No := 5,   // "Safety_Stops_FB"
                    Mode := "Control_DB".VTD_Sys[5].Mode,
                    Timeout := "Settings_DB".LCnv_Sys[5].Cnv_Level[1].Cnv1.Safety_stop_Timeout,
                    Reset := "Control_DB".LCnv_Sys[5].Cnv_Level[1].Cnv1.Instruction.Reset,
                    Sfts_Control := "Control_DB".LCnv_Sys[5].Cnv_Level[1].Cnv1.Safety_Stop_Cnrl,
                    ENO => #_w1);
   "Sf_C5102_FB_DB"(EN := #_w1,   // "Safety_Stops_FB"
                    Sys_No := 5,
                    Mode := "Control_DB".VTD_Sys[5].Mode,
                    Timeout := "Settings_DB".LCnv_Sys[5].Cnv_Level[2].Cnv1.Safety_stop_Timeout,
                    Reset := "Control_DB".LCnv_Sys[5].Cnv_Level[2].Cnv1.Instruction.Reset,
                    Sfts_Control := "Control_DB".LCnv_Sys[5].Cnv_Level[2].Cnv1.Safety_Stop_Cnrl,
                    ENO => #_w2);
   IF #_w2 THEN
       "Sf_C5103_FB_DB"(Sys_No := 5,   // "Safety_Stops_FB"
                        Mode := "Control_DB".VTD_Sys[5].Mode,
                        Timeout := "Settings_DB".LCnv_Sys[5].Cnv_Level[3].Cnv1.Safety_stop_Timeout,
                        Reset := "Control_DB".LCnv_Sys[5].Cnv_Level[3].Cnv1.Instruction.Reset,
                        Sfts_Control := "Control_DB".LCnv_Sys[5].Cnv_Level[3].Cnv1.Safety_Stop_Cnrl);
   END_IF;
   "Sf_C5104_FB_DB"(Sys_No := 5,   // "Safety_Stops_FB"
                    Mode := "Control_DB".VTD_Sys[5].Mode,
                    Timeout := "Settings_DB".LCnv_Sys[5].Cnv_Level[4].Cnv1.Safety_stop_Timeout,
                    Reset := "Control_DB".LCnv_Sys[5].Cnv_Level[4].Cnv1.Instruction.Reset,
                    Sfts_Control := "Control_DB".LCnv_Sys[5].Cnv_Level[4].Cnv1.Safety_Stop_Cnrl,
                    ENO => #_w3);
   "Sf_C5105_FB_DB"(EN := #_w3,   // "Safety_Stops_FB"
                    Sys_No := 5,
                    Mode := "Control_DB".VTD_Sys[5].Mode,
                    Timeout := "Settings_DB".LCnv_Sys[5].Cnv_Level[5].Cnv1.Safety_stop_Timeout,
                    Reset := "Control_DB".LCnv_Sys[5].Cnv_Level[5].Cnv1.Instruction.Reset,
                    Sfts_Control := "Control_DB".LCnv_Sys[5].Cnv_Level[5].Cnv1.Safety_Stop_Cnrl,
                    ENO => #_w4);
   IF #_w4 THEN
       "Sf_C5106_FB_DB"(Sys_No := 5,   // "Safety_Stops_FB"
                        Mode := "Control_DB".VTD_Sys[5].Mode,
                        Timeout := "Settings_DB".LCnv_Sys[5].Cnv_Level[6].Cnv1.Safety_stop_Timeout,
                        Reset := "Control_DB".LCnv_Sys[5].Cnv_Level[6].Cnv1.Instruction.Reset,
                        Sfts_Control := "Control_DB".LCnv_Sys[5].Cnv_Level[6].Cnv1.Safety_Stop_Cnrl);
   END_IF;
   "Sf_C5107_FB_DB"(Sys_No := 5,   // "Safety_Stops_FB"
                    Mode := "Control_DB".VTD_Sys[5].Mode,
                    Timeout := "Settings_DB".LCnv_Sys[5].Cnv_Level[7].Cnv1.Safety_stop_Timeout,
                    Reset := "Control_DB".LCnv_Sys[5].Cnv_Level[7].Cnv1.Instruction.Reset,
                    Sfts_Control := "Control_DB".LCnv_Sys[5].Cnv_Level[7].Cnv1.Safety_Stop_Cnrl,
                    ENO => #_w5);
   IF #_w5 THEN
       "Sf_C5108_FB_DB"(Sys_No := 5,   // "Safety_Stops_FB"
                        Mode := "Control_DB".VTD_Sys[5].Mode,
                        Timeout := "Settings_DB".LCnv_Sys[5].Cnv_Level[8].Cnv1.Safety_stop_Timeout,
                        Reset := "Control_DB".LCnv_Sys[5].Cnv_Level[8].Cnv1.Instruction.Reset,
                        Sfts_Control := "Control_DB".LCnv_Sys[5].Cnv_Level[8].Cnv1.Safety_Stop_Cnrl);
   END_IF;
END_REGION

REGION Network 40: Light bars
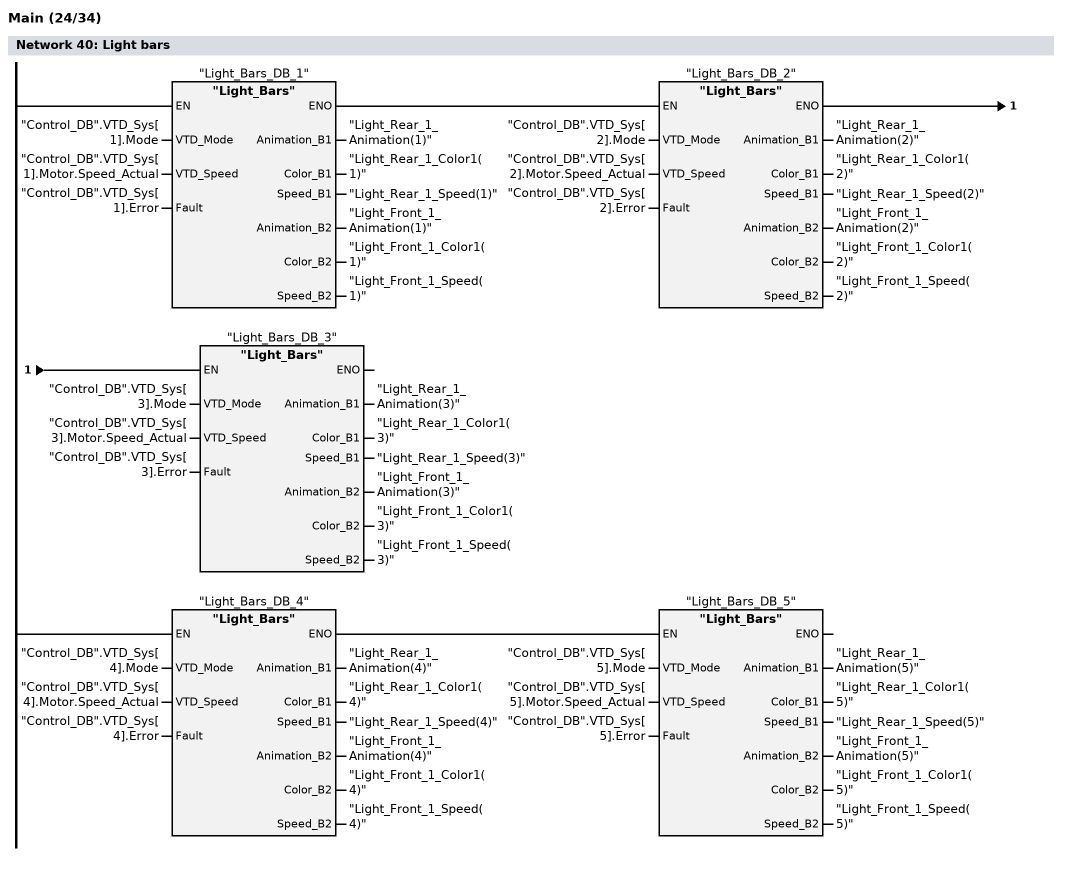
   RUNG wire#powerrail
      "Light_Bars_DB_1"(VTD_Mode := "Control_DB".VTD_Sys[1].Mode, VTD_Speed := "Control_DB".VTD_Sys[1].Motor.Speed_Actual, Fault := "Control_DB".VTD_Sys[1].Error, Animation_B1 => "Light_Rear_1_Animation(1)", Color_B1 => "Light_Rear_1_Color1(1)", Speed_B1 => "Light_Rear_1_Speed(1)", Animation_B2 => "Light_Front_1_Animation(1)", Color_B2 => "Light_Front_1_Color1(1)", Speed_B2 => "Light_Front_1_Speed(1)")
      "Light_Bars_DB_2"(VTD_Mode := "Control_DB".VTD_Sys[2].Mode, VTD_Speed := "Control_DB".VTD_Sys[2].Motor.Speed_Actual, Fault := "Control_DB".VTD_Sys[2].Error, Animation_B1 => "Light_Rear_1_Animation(2)", Color_B1 => "Light_Rear_1_Color1(2)", Speed_B1 => "Light_Rear_1_Speed(2)", Animation_B2 => "Light_Front_1_Animation(2)", Color_B2 => "Light_Front_1_Color1(2)", Speed_B2 => "Light_Front_1_Speed(2)")
      "Light_Bars_DB_3"(VTD_Mode := "Control_DB".VTD_Sys[3].Mode, VTD_Speed := "Control_DB".VTD_Sys[3].Motor.Speed_Actual, Fault := "Control_DB".VTD_Sys[3].Error, Animation_B1 => "Light_Rear_1_Animation(3)", Color_B1 => "Light_Rear_1_Color1(3)", Speed_B1 => "Light_Rear_1_Speed(3)", Animation_B2 => "Light_Front_1_Animation(3)", Color_B2 => "Light_Front_1_Color1(3)", Speed_B2 => "Light_Front_1_Speed(3)")
   END_RUNG
   RUNG wire#powerrail
      "Light_Bars_DB_4"(VTD_Mode := "Control_DB".VTD_Sys[4].Mode, VTD_Speed := "Control_DB".VTD_Sys[4].Motor.Speed_Actual, Fault := "Control_DB".VTD_Sys[4].Error, Animation_B1 => "Light_Rear_1_Animation(4)", Color_B1 => "Light_Rear_1_Color1(4)", Speed_B1 => "Light_Rear_1_Speed(4)", Animation_B2 => "Light_Front_1_Animation(4)", Color_B2 => "Light_Front_1_Color1(4)", Speed_B2 => "Light_Front_1_Speed(4)")
      "Light_Bars_DB_5"(VTD_Mode := "Control_DB".VTD_Sys[5].Mode, VTD_Speed := "Control_DB".VTD_Sys[5].Motor.Speed_Actual, Fault := "Control_DB".VTD_Sys[5].Error, Animation_B1 => "Light_Rear_1_Animation(5)", Color_B1 => "Light_Rear_1_Color1(5)", Speed_B1 => "Light_Rear_1_Speed(5)", Animation_B2 => "Light_Front_1_Animation(5)", Color_B2 => "Light_Front_1_Color1(5)", Speed_B2 => "Light_Front_1_Speed(5)")
   END_RUNG
   // the same network as SCL:
   "Light_Bars_DB_1"(VTD_Mode := "Control_DB".VTD_Sys[1].Mode,   // "Light_Bars"
                     VTD_Speed := "Control_DB".VTD_Sys[1].Motor.Speed_Actual,
                     Fault := "Control_DB".VTD_Sys[1].Error,
                     Animation_B1 => "Light_Rear_1_Animation(1)",
                     Color_B1 => "Light_Rear_1_Color1(1)",
                     Speed_B1 => "Light_Rear_1_Speed(1)",
                     Animation_B2 => "Light_Front_1_Animation(1)",
                     Color_B2 => "Light_Front_1_Color1(1)",
                     Speed_B2 => "Light_Front_1_Speed(1)",
                     ENO => #_w1);
   "Light_Bars_DB_2"(EN := #_w1,   // "Light_Bars"
                     VTD_Mode := "Control_DB".VTD_Sys[2].Mode,
                     VTD_Speed := "Control_DB".VTD_Sys[2].Motor.Speed_Actual,
                     Fault := "Control_DB".VTD_Sys[2].Error,
                     Animation_B1 => "Light_Rear_1_Animation(2)",
                     Color_B1 => "Light_Rear_1_Color1(2)",
                     Speed_B1 => "Light_Rear_1_Speed(2)",
                     Animation_B2 => "Light_Front_1_Animation(2)",
                     Color_B2 => "Light_Front_1_Color1(2)",
                     Speed_B2 => "Light_Front_1_Speed(2)",
                     ENO => #_w2);
   IF #_w2 THEN
       "Light_Bars_DB_3"(VTD_Mode := "Control_DB".VTD_Sys[3].Mode,   // "Light_Bars"
                         VTD_Speed := "Control_DB".VTD_Sys[3].Motor.Speed_Actual,
                         Fault := "Control_DB".VTD_Sys[3].Error,
                         Animation_B1 => "Light_Rear_1_Animation(3)",
                         Color_B1 => "Light_Rear_1_Color1(3)",
                         Speed_B1 => "Light_Rear_1_Speed(3)",
                         Animation_B2 => "Light_Front_1_Animation(3)",
                         Color_B2 => "Light_Front_1_Color1(3)",
                         Speed_B2 => "Light_Front_1_Speed(3)");
   END_IF;
   "Light_Bars_DB_4"(VTD_Mode := "Control_DB".VTD_Sys[4].Mode,   // "Light_Bars"
                     VTD_Speed := "Control_DB".VTD_Sys[4].Motor.Speed_Actual,
                     Fault := "Control_DB".VTD_Sys[4].Error,
                     Animation_B1 => "Light_Rear_1_Animation(4)",
                     Color_B1 => "Light_Rear_1_Color1(4)",
                     Speed_B1 => "Light_Rear_1_Speed(4)",
                     Animation_B2 => "Light_Front_1_Animation(4)",
                     Color_B2 => "Light_Front_1_Color1(4)",
                     Speed_B2 => "Light_Front_1_Speed(4)",
                     ENO => #_w3);
   IF #_w3 THEN
       "Light_Bars_DB_5"(VTD_Mode := "Control_DB".VTD_Sys[5].Mode,   // "Light_Bars"
                         VTD_Speed := "Control_DB".VTD_Sys[5].Motor.Speed_Actual,
                         Fault := "Control_DB".VTD_Sys[5].Error,
                         Animation_B1 => "Light_Rear_1_Animation(5)",
                         Color_B1 => "Light_Rear_1_Color1(5)",
                         Speed_B1 => "Light_Rear_1_Speed(5)",
                         Animation_B2 => "Light_Front_1_Animation(5)",
                         Color_B2 => "Light_Front_1_Color1(5)",
                         Speed_B2 => "Light_Front_1_Speed(5)");
   END_IF;
END_REGION

REGION Network 41: Barcode - System 1
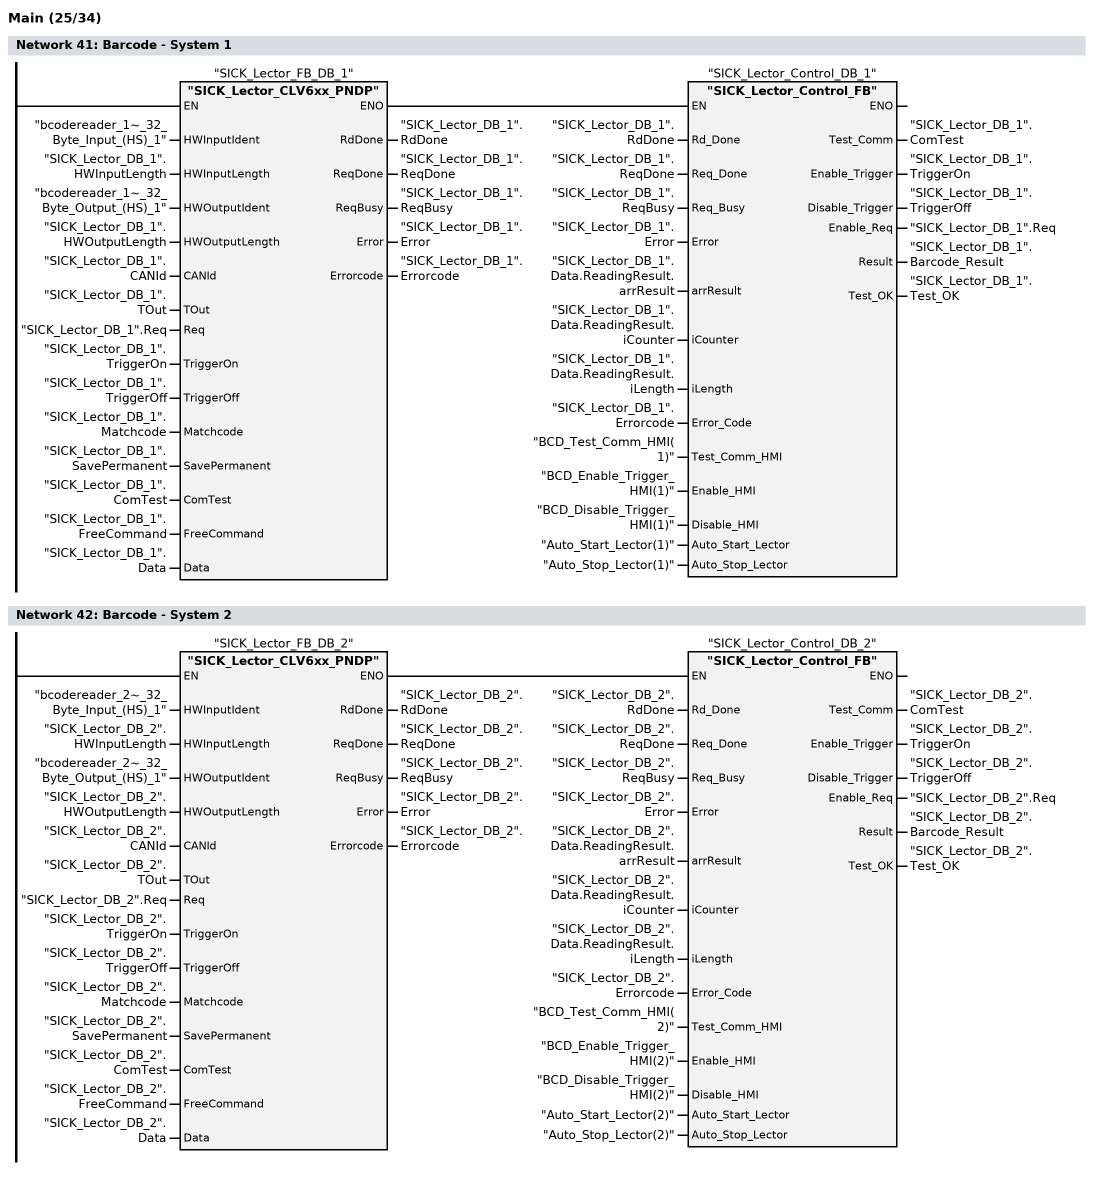
   RUNG wire#powerrail
      "SICK_Lector_FB_DB_1"(HWInputIdent := "bcodereader_1~_32_Byte_Input_(HS)_1", HWInputLength := "SICK_Lector_DB_1".HWInputLength, HWOutputIdent := "bcodereader_1~_32_Byte_Output_(HS)_1", HWOutputLength := "SICK_Lector_DB_1".HWOutputLength, CANId := "SICK_Lector_DB_1".CANId, TOut := "SICK_Lector_DB_1".TOut, Req := "SICK_Lector_DB_1".Req, TriggerOn := "SICK_Lector_DB_1".TriggerOn, TriggerOff := "SICK_Lector_DB_1".TriggerOff, Matchcode := "SICK_Lector_DB_1".Matchcode, SavePermanent := "SICK_Lector_DB_1".SavePermanent, ComTest := "SICK_Lector_DB_1".ComTest, FreeCommand := "SICK_Lector_DB_1".FreeCommand, Data := "SICK_Lector_DB_1".Data, RdDone => "SICK_Lector_DB_1".RdDone, ReqDone => "SICK_Lector_DB_1".ReqDone, ReqBusy => "SICK_Lector_DB_1".ReqBusy, Error => "SICK_Lector_DB_1".Error, Errorcode => "SICK_Lector_DB_1".Errorcode)
      "SICK_Lector_Control_DB_1"(Rd_Done := "SICK_Lector_DB_1".RdDone, Req_Done := "SICK_Lector_DB_1".ReqDone, Req_Busy := "SICK_Lector_DB_1".ReqBusy, Error := "SICK_Lector_DB_1".Error, arrResult := "SICK_Lector_DB_1".Data.ReadingResult.arrResult, iCounter := "SICK_Lector_DB_1".Data.ReadingResult.iCounter, iLength := "SICK_Lector_DB_1".Data.ReadingResult.iLength, Error_Code := "SICK_Lector_DB_1".Errorcode, Test_Comm_HMI := "BCD_Test_Comm_HMI(1)", Enable_HMI := "BCD_Enable_Trigger_HMI(1)", Disable_HMI := "BCD_Disable_Trigger_HMI(1)", Auto_Start_Lector := "Auto_Start_Lector(1)", Auto_Stop_Lector := "Auto_Stop_Lector(1)", Test_Comm => "SICK_Lector_DB_1".ComTest, Enable_Trigger => "SICK_Lector_DB_1".TriggerOn, Disable_Trigger => "SICK_Lector_DB_1".TriggerOff, Enable_Req => "SICK_Lector_DB_1".Req, Result => "SICK_Lector_DB_1".Barcode_Result, Test_OK => "SICK_Lector_DB_1".Test_OK)
   END_RUNG
   // the same network as SCL:
   "SICK_Lector_FB_DB_1"(HWInputIdent := "bcodereader_1~_32_Byte_Input_(HS)_1",   // "SICK_Lector_CLV6xx_PNDP"
                         HWInputLength := "SICK_Lector_DB_1".HWInputLength,
                         HWOutputIdent := "bcodereader_1~_32_Byte_Output_(HS)_1",
                         HWOutputLength := "SICK_Lector_DB_1".HWOutputLength,
                         CANId := "SICK_Lector_DB_1".CANId,
                         TOut := "SICK_Lector_DB_1".TOut,
                         Req := "SICK_Lector_DB_1".Req,
                         TriggerOn := "SICK_Lector_DB_1".TriggerOn,
                         TriggerOff := "SICK_Lector_DB_1".TriggerOff,
                         Matchcode := "SICK_Lector_DB_1".Matchcode,
                         SavePermanent := "SICK_Lector_DB_1".SavePermanent,
                         ComTest := "SICK_Lector_DB_1".ComTest,
                         FreeCommand := "SICK_Lector_DB_1".FreeCommand,
                         Data := "SICK_Lector_DB_1".Data,
                         RdDone => "SICK_Lector_DB_1".RdDone,
                         ReqDone => "SICK_Lector_DB_1".ReqDone,
                         ReqBusy => "SICK_Lector_DB_1".ReqBusy,
                         Error => "SICK_Lector_DB_1".Error,
                         Errorcode => "SICK_Lector_DB_1".Errorcode,
                         ENO => #_w1);
   IF #_w1 THEN
       "SICK_Lector_Control_DB_1"(Rd_Done := "SICK_Lector_DB_1".RdDone,   // "SICK_Lector_Control_FB"
                               Req_Done := "SICK_Lector_DB_1".ReqDone,
                               Req_Busy := "SICK_Lector_DB_1".ReqBusy,
                               Error := "SICK_Lector_DB_1".Error,
                               arrResult := "SICK_Lector_DB_1".Data.ReadingResult.arrResult,
                               iCounter := "SICK_Lector_DB_1".Data.ReadingResult.iCounter,
                               iLength := "SICK_Lector_DB_1".Data.ReadingResult.iLength,
                               Error_Code := "SICK_Lector_DB_1".Errorcode,
                               Test_Comm_HMI := "BCD_Test_Comm_HMI(1)",
                               Enable_HMI := "BCD_Enable_Trigger_HMI(1)",
                               Disable_HMI := "BCD_Disable_Trigger_HMI(1)",
                               Auto_Start_Lector := "Auto_Start_Lector(1)",
                               Auto_Stop_Lector := "Auto_Stop_Lector(1)",
                               Test_Comm => "SICK_Lector_DB_1".ComTest,
                               Enable_Trigger => "SICK_Lector_DB_1".TriggerOn,
                               Disable_Trigger => "SICK_Lector_DB_1".TriggerOff,
                               Enable_Req => "SICK_Lector_DB_1".Req,
                               Result => "SICK_Lector_DB_1".Barcode_Result,
                               Test_OK => "SICK_Lector_DB_1".Test_OK);
   END_IF;
END_REGION

REGION Network 42: Barcode - System 2
   RUNG wire#powerrail
      "SICK_Lector_FB_DB_2"(HWInputIdent := "bcodereader_2~_32_Byte_Input_(HS)_1", HWInputLength := "SICK_Lector_DB_2".HWInputLength, HWOutputIdent := "bcodereader_2~_32_Byte_Output_(HS)_1", HWOutputLength := "SICK_Lector_DB_2".HWOutputLength, CANId := "SICK_Lector_DB_2".CANId, TOut := "SICK_Lector_DB_2".TOut, Req := "SICK_Lector_DB_2".Req, TriggerOn := "SICK_Lector_DB_2".TriggerOn, TriggerOff := "SICK_Lector_DB_2".TriggerOff, Matchcode := "SICK_Lector_DB_2".Matchcode, SavePermanent := "SICK_Lector_DB_2".SavePermanent, ComTest := "SICK_Lector_DB_2".ComTest, FreeCommand := "SICK_Lector_DB_2".FreeCommand, Data := "SICK_Lector_DB_2".Data, RdDone => "SICK_Lector_DB_2".RdDone, ReqDone => "SICK_Lector_DB_2".ReqDone, ReqBusy => "SICK_Lector_DB_2".ReqBusy, Error => "SICK_Lector_DB_2".Error, Errorcode => "SICK_Lector_DB_2".Errorcode)
      "SICK_Lector_Control_DB_2"(Rd_Done := "SICK_Lector_DB_2".RdDone, Req_Done := "SICK_Lector_DB_2".ReqDone, Req_Busy := "SICK_Lector_DB_2".ReqBusy, Error := "SICK_Lector_DB_2".Error, arrResult := "SICK_Lector_DB_2".Data.ReadingResult.arrResult, iCounter := "SICK_Lector_DB_2".Data.ReadingResult.iCounter, iLength := "SICK_Lector_DB_2".Data.ReadingResult.iLength, Error_Code := "SICK_Lector_DB_2".Errorcode, Test_Comm_HMI := "BCD_Test_Comm_HMI(2)", Enable_HMI := "BCD_Enable_Trigger_HMI(2)", Disable_HMI := "BCD_Disable_Trigger_HMI(2)", Auto_Start_Lector := "Auto_Start_Lector(2)", Auto_Stop_Lector := "Auto_Stop_Lector(2)", Test_Comm => "SICK_Lector_DB_2".ComTest, Enable_Trigger => "SICK_Lector_DB_2".TriggerOn, Disable_Trigger => "SICK_Lector_DB_2".TriggerOff, Enable_Req => "SICK_Lector_DB_2".Req, Result => "SICK_Lector_DB_2".Barcode_Result, Test_OK => "SICK_Lector_DB_2".Test_OK)
   END_RUNG
   // the same network as SCL:
   "SICK_Lector_FB_DB_2"(HWInputIdent := "bcodereader_2~_32_Byte_Input_(HS)_1",   // "SICK_Lector_CLV6xx_PNDP"
                         HWInputLength := "SICK_Lector_DB_2".HWInputLength,
                         HWOutputIdent := "bcodereader_2~_32_Byte_Output_(HS)_1",
                         HWOutputLength := "SICK_Lector_DB_2".HWOutputLength,
                         CANId := "SICK_Lector_DB_2".CANId,
                         TOut := "SICK_Lector_DB_2".TOut,
                         Req := "SICK_Lector_DB_2".Req,
                         TriggerOn := "SICK_Lector_DB_2".TriggerOn,
                         TriggerOff := "SICK_Lector_DB_2".TriggerOff,
                         Matchcode := "SICK_Lector_DB_2".Matchcode,
                         SavePermanent := "SICK_Lector_DB_2".SavePermanent,
                         ComTest := "SICK_Lector_DB_2".ComTest,
                         FreeCommand := "SICK_Lector_DB_2".FreeCommand,
                         Data := "SICK_Lector_DB_2".Data,
                         RdDone => "SICK_Lector_DB_2".RdDone,
                         ReqDone => "SICK_Lector_DB_2".ReqDone,
                         ReqBusy => "SICK_Lector_DB_2".ReqBusy,
                         Error => "SICK_Lector_DB_2".Error,
                         Errorcode => "SICK_Lector_DB_2".Errorcode,
                         ENO => #_w1);
   IF #_w1 THEN
       "SICK_Lector_Control_DB_2"(Rd_Done := "SICK_Lector_DB_2".RdDone,   // "SICK_Lector_Control_FB"
                               Req_Done := "SICK_Lector_DB_2".ReqDone,
                               Req_Busy := "SICK_Lector_DB_2".ReqBusy,
                               Error := "SICK_Lector_DB_2".Error,
                               arrResult := "SICK_Lector_DB_2".Data.ReadingResult.arrResult,
                               iCounter := "SICK_Lector_DB_2".Data.ReadingResult.iCounter,
                               iLength := "SICK_Lector_DB_2".Data.ReadingResult.iLength,
                               Error_Code := "SICK_Lector_DB_2".Errorcode,
                               Test_Comm_HMI := "BCD_Test_Comm_HMI(2)",
                               Enable_HMI := "BCD_Enable_Trigger_HMI(2)",
                               Disable_HMI := "BCD_Disable_Trigger_HMI(2)",
                               Auto_Start_Lector := "Auto_Start_Lector(2)",
                               Auto_Stop_Lector := "Auto_Stop_Lector(2)",
                               Test_Comm => "SICK_Lector_DB_2".ComTest,
                               Enable_Trigger => "SICK_Lector_DB_2".TriggerOn,
                               Disable_Trigger => "SICK_Lector_DB_2".TriggerOff,
                               Enable_Req => "SICK_Lector_DB_2".Req,
                               Result => "SICK_Lector_DB_2".Barcode_Result,
                               Test_OK => "SICK_Lector_DB_2".Test_OK);
   END_IF;
END_REGION

REGION Network 43: Barcode - System 3
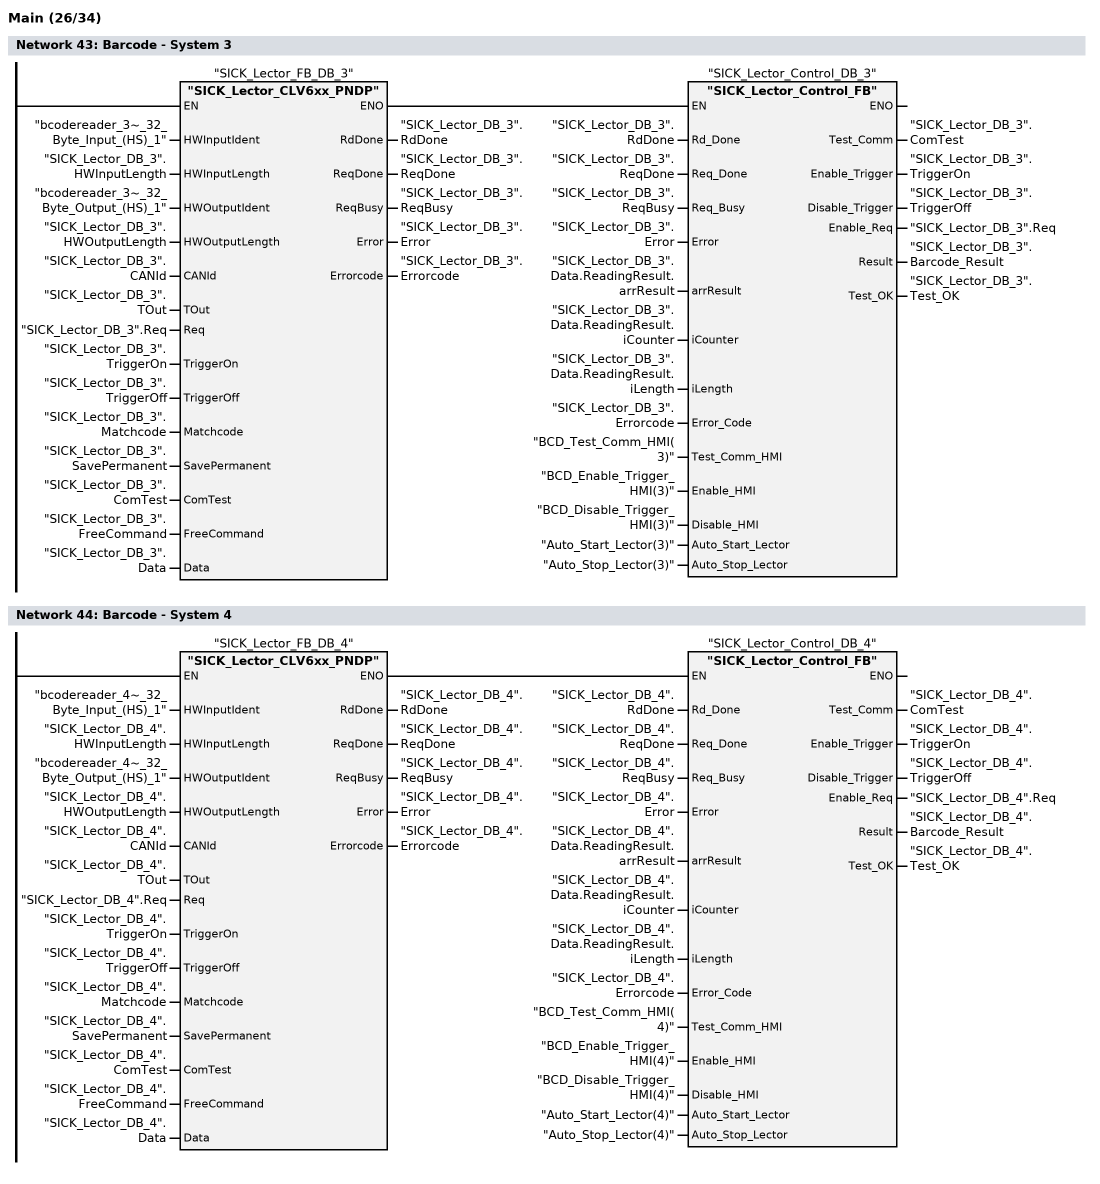
   RUNG wire#powerrail
      "SICK_Lector_FB_DB_3"(HWInputIdent := "bcodereader_3~_32_Byte_Input_(HS)_1", HWInputLength := "SICK_Lector_DB_3".HWInputLength, HWOutputIdent := "bcodereader_3~_32_Byte_Output_(HS)_1", HWOutputLength := "SICK_Lector_DB_3".HWOutputLength, CANId := "SICK_Lector_DB_3".CANId, TOut := "SICK_Lector_DB_3".TOut, Req := "SICK_Lector_DB_3".Req, TriggerOn := "SICK_Lector_DB_3".TriggerOn, TriggerOff := "SICK_Lector_DB_3".TriggerOff, Matchcode := "SICK_Lector_DB_3".Matchcode, SavePermanent := "SICK_Lector_DB_3".SavePermanent, ComTest := "SICK_Lector_DB_3".ComTest, FreeCommand := "SICK_Lector_DB_3".FreeCommand, Data := "SICK_Lector_DB_3".Data, RdDone => "SICK_Lector_DB_3".RdDone, ReqDone => "SICK_Lector_DB_3".ReqDone, ReqBusy => "SICK_Lector_DB_3".ReqBusy, Error => "SICK_Lector_DB_3".Error, Errorcode => "SICK_Lector_DB_3".Errorcode)
      "SICK_Lector_Control_DB_3"(Rd_Done := "SICK_Lector_DB_3".RdDone, Req_Done := "SICK_Lector_DB_3".ReqDone, Req_Busy := "SICK_Lector_DB_3".ReqBusy, Error := "SICK_Lector_DB_3".Error, arrResult := "SICK_Lector_DB_3".Data.ReadingResult.arrResult, iCounter := "SICK_Lector_DB_3".Data.ReadingResult.iCounter, iLength := "SICK_Lector_DB_3".Data.ReadingResult.iLength, Error_Code := "SICK_Lector_DB_3".Errorcode, Test_Comm_HMI := "BCD_Test_Comm_HMI(3)", Enable_HMI := "BCD_Enable_Trigger_HMI(3)", Disable_HMI := "BCD_Disable_Trigger_HMI(3)", Auto_Start_Lector := "Auto_Start_Lector(3)", Auto_Stop_Lector := "Auto_Stop_Lector(3)", Test_Comm => "SICK_Lector_DB_3".ComTest, Enable_Trigger => "SICK_Lector_DB_3".TriggerOn, Disable_Trigger => "SICK_Lector_DB_3".TriggerOff, Enable_Req => "SICK_Lector_DB_3".Req, Result => "SICK_Lector_DB_3".Barcode_Result, Test_OK => "SICK_Lector_DB_3".Test_OK)
   END_RUNG
   // the same network as SCL:
   "SICK_Lector_FB_DB_3"(HWInputIdent := "bcodereader_3~_32_Byte_Input_(HS)_1",   // "SICK_Lector_CLV6xx_PNDP"
                         HWInputLength := "SICK_Lector_DB_3".HWInputLength,
                         HWOutputIdent := "bcodereader_3~_32_Byte_Output_(HS)_1",
                         HWOutputLength := "SICK_Lector_DB_3".HWOutputLength,
                         CANId := "SICK_Lector_DB_3".CANId,
                         TOut := "SICK_Lector_DB_3".TOut,
                         Req := "SICK_Lector_DB_3".Req,
                         TriggerOn := "SICK_Lector_DB_3".TriggerOn,
                         TriggerOff := "SICK_Lector_DB_3".TriggerOff,
                         Matchcode := "SICK_Lector_DB_3".Matchcode,
                         SavePermanent := "SICK_Lector_DB_3".SavePermanent,
                         ComTest := "SICK_Lector_DB_3".ComTest,
                         FreeCommand := "SICK_Lector_DB_3".FreeCommand,
                         Data := "SICK_Lector_DB_3".Data,
                         RdDone => "SICK_Lector_DB_3".RdDone,
                         ReqDone => "SICK_Lector_DB_3".ReqDone,
                         ReqBusy => "SICK_Lector_DB_3".ReqBusy,
                         Error => "SICK_Lector_DB_3".Error,
                         Errorcode => "SICK_Lector_DB_3".Errorcode,
                         ENO => #_w1);
   IF #_w1 THEN
       "SICK_Lector_Control_DB_3"(Rd_Done := "SICK_Lector_DB_3".RdDone,   // "SICK_Lector_Control_FB"
                               Req_Done := "SICK_Lector_DB_3".ReqDone,
                               Req_Busy := "SICK_Lector_DB_3".ReqBusy,
                               Error := "SICK_Lector_DB_3".Error,
                               arrResult := "SICK_Lector_DB_3".Data.ReadingResult.arrResult,
                               iCounter := "SICK_Lector_DB_3".Data.ReadingResult.iCounter,
                               iLength := "SICK_Lector_DB_3".Data.ReadingResult.iLength,
                               Error_Code := "SICK_Lector_DB_3".Errorcode,
                               Test_Comm_HMI := "BCD_Test_Comm_HMI(3)",
                               Enable_HMI := "BCD_Enable_Trigger_HMI(3)",
                               Disable_HMI := "BCD_Disable_Trigger_HMI(3)",
                               Auto_Start_Lector := "Auto_Start_Lector(3)",
                               Auto_Stop_Lector := "Auto_Stop_Lector(3)",
                               Test_Comm => "SICK_Lector_DB_3".ComTest,
                               Enable_Trigger => "SICK_Lector_DB_3".TriggerOn,
                               Disable_Trigger => "SICK_Lector_DB_3".TriggerOff,
                               Enable_Req => "SICK_Lector_DB_3".Req,
                               Result => "SICK_Lector_DB_3".Barcode_Result,
                               Test_OK => "SICK_Lector_DB_3".Test_OK);
   END_IF;
END_REGION

REGION Network 44: Barcode - System 4
   RUNG wire#powerrail
      "SICK_Lector_FB_DB_4"(HWInputIdent := "bcodereader_4~_32_Byte_Input_(HS)_1", HWInputLength := "SICK_Lector_DB_4".HWInputLength, HWOutputIdent := "bcodereader_4~_32_Byte_Output_(HS)_1", HWOutputLength := "SICK_Lector_DB_4".HWOutputLength, CANId := "SICK_Lector_DB_4".CANId, TOut := "SICK_Lector_DB_4".TOut, Req := "SICK_Lector_DB_4".Req, TriggerOn := "SICK_Lector_DB_4".TriggerOn, TriggerOff := "SICK_Lector_DB_4".TriggerOff, Matchcode := "SICK_Lector_DB_4".Matchcode, SavePermanent := "SICK_Lector_DB_4".SavePermanent, ComTest := "SICK_Lector_DB_4".ComTest, FreeCommand := "SICK_Lector_DB_4".FreeCommand, Data := "SICK_Lector_DB_4".Data, RdDone => "SICK_Lector_DB_4".RdDone, ReqDone => "SICK_Lector_DB_4".ReqDone, ReqBusy => "SICK_Lector_DB_4".ReqBusy, Error => "SICK_Lector_DB_4".Error, Errorcode => "SICK_Lector_DB_4".Errorcode)
      "SICK_Lector_Control_DB_4"(Rd_Done := "SICK_Lector_DB_4".RdDone, Req_Done := "SICK_Lector_DB_4".ReqDone, Req_Busy := "SICK_Lector_DB_4".ReqBusy, Error := "SICK_Lector_DB_4".Error, arrResult := "SICK_Lector_DB_4".Data.ReadingResult.arrResult, iCounter := "SICK_Lector_DB_4".Data.ReadingResult.iCounter, iLength := "SICK_Lector_DB_4".Data.ReadingResult.iLength, Error_Code := "SICK_Lector_DB_4".Errorcode, Test_Comm_HMI := "BCD_Test_Comm_HMI(4)", Enable_HMI := "BCD_Enable_Trigger_HMI(4)", Disable_HMI := "BCD_Disable_Trigger_HMI(4)", Auto_Start_Lector := "Auto_Start_Lector(4)", Auto_Stop_Lector := "Auto_Stop_Lector(4)", Test_Comm => "SICK_Lector_DB_4".ComTest, Enable_Trigger => "SICK_Lector_DB_4".TriggerOn, Disable_Trigger => "SICK_Lector_DB_4".TriggerOff, Enable_Req => "SICK_Lector_DB_4".Req, Result => "SICK_Lector_DB_4".Barcode_Result, Test_OK => "SICK_Lector_DB_4".Test_OK)
   END_RUNG
   // the same network as SCL:
   "SICK_Lector_FB_DB_4"(HWInputIdent := "bcodereader_4~_32_Byte_Input_(HS)_1",   // "SICK_Lector_CLV6xx_PNDP"
                         HWInputLength := "SICK_Lector_DB_4".HWInputLength,
                         HWOutputIdent := "bcodereader_4~_32_Byte_Output_(HS)_1",
                         HWOutputLength := "SICK_Lector_DB_4".HWOutputLength,
                         CANId := "SICK_Lector_DB_4".CANId,
                         TOut := "SICK_Lector_DB_4".TOut,
                         Req := "SICK_Lector_DB_4".Req,
                         TriggerOn := "SICK_Lector_DB_4".TriggerOn,
                         TriggerOff := "SICK_Lector_DB_4".TriggerOff,
                         Matchcode := "SICK_Lector_DB_4".Matchcode,
                         SavePermanent := "SICK_Lector_DB_4".SavePermanent,
                         ComTest := "SICK_Lector_DB_4".ComTest,
                         FreeCommand := "SICK_Lector_DB_4".FreeCommand,
                         Data := "SICK_Lector_DB_4".Data,
                         RdDone => "SICK_Lector_DB_4".RdDone,
                         ReqDone => "SICK_Lector_DB_4".ReqDone,
                         ReqBusy => "SICK_Lector_DB_4".ReqBusy,
                         Error => "SICK_Lector_DB_4".Error,
                         Errorcode => "SICK_Lector_DB_4".Errorcode,
                         ENO => #_w1);
   IF #_w1 THEN
       "SICK_Lector_Control_DB_4"(Rd_Done := "SICK_Lector_DB_4".RdDone,   // "SICK_Lector_Control_FB"
                               Req_Done := "SICK_Lector_DB_4".ReqDone,
                               Req_Busy := "SICK_Lector_DB_4".ReqBusy,
                               Error := "SICK_Lector_DB_4".Error,
                               arrResult := "SICK_Lector_DB_4".Data.ReadingResult.arrResult,
                               iCounter := "SICK_Lector_DB_4".Data.ReadingResult.iCounter,
                               iLength := "SICK_Lector_DB_4".Data.ReadingResult.iLength,
                               Error_Code := "SICK_Lector_DB_4".Errorcode,
                               Test_Comm_HMI := "BCD_Test_Comm_HMI(4)",
                               Enable_HMI := "BCD_Enable_Trigger_HMI(4)",
                               Disable_HMI := "BCD_Disable_Trigger_HMI(4)",
                               Auto_Start_Lector := "Auto_Start_Lector(4)",
                               Auto_Stop_Lector := "Auto_Stop_Lector(4)",
                               Test_Comm => "SICK_Lector_DB_4".ComTest,
                               Enable_Trigger => "SICK_Lector_DB_4".TriggerOn,
                               Disable_Trigger => "SICK_Lector_DB_4".TriggerOff,
                               Enable_Req => "SICK_Lector_DB_4".Req,
                               Result => "SICK_Lector_DB_4".Barcode_Result,
                               Test_OK => "SICK_Lector_DB_4".Test_OK);
   END_IF;
END_REGION

REGION Network 45: Barcode - System 5
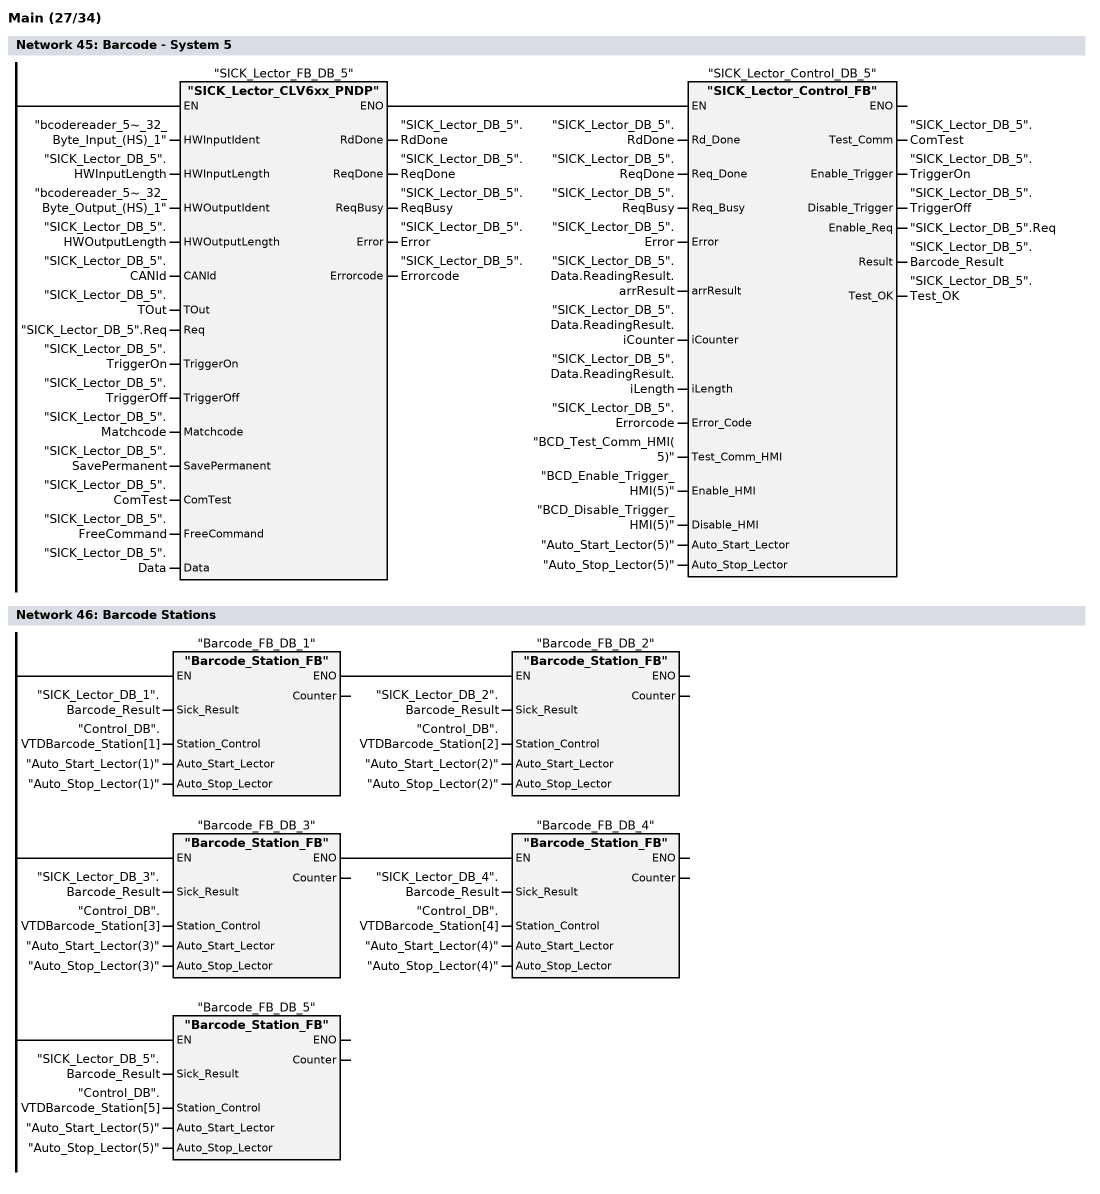
   RUNG wire#powerrail
      "SICK_Lector_FB_DB_5"(HWInputIdent := "bcodereader_5~_32_Byte_Input_(HS)_1", HWInputLength := "SICK_Lector_DB_5".HWInputLength, HWOutputIdent := "bcodereader_5~_32_Byte_Output_(HS)_1", HWOutputLength := "SICK_Lector_DB_5".HWOutputLength, CANId := "SICK_Lector_DB_5".CANId, TOut := "SICK_Lector_DB_5".TOut, Req := "SICK_Lector_DB_5".Req, TriggerOn := "SICK_Lector_DB_5".TriggerOn, TriggerOff := "SICK_Lector_DB_5".TriggerOff, Matchcode := "SICK_Lector_DB_5".Matchcode, SavePermanent := "SICK_Lector_DB_5".SavePermanent, ComTest := "SICK_Lector_DB_5".ComTest, FreeCommand := "SICK_Lector_DB_5".FreeCommand, Data := "SICK_Lector_DB_5".Data, RdDone => "SICK_Lector_DB_5".RdDone, ReqDone => "SICK_Lector_DB_5".ReqDone, ReqBusy => "SICK_Lector_DB_5".ReqBusy, Error => "SICK_Lector_DB_5".Error, Errorcode => "SICK_Lector_DB_5".Errorcode)
      "SICK_Lector_Control_DB_5"(Rd_Done := "SICK_Lector_DB_5".RdDone, Req_Done := "SICK_Lector_DB_5".ReqDone, Req_Busy := "SICK_Lector_DB_5".ReqBusy, Error := "SICK_Lector_DB_5".Error, arrResult := "SICK_Lector_DB_5".Data.ReadingResult.arrResult, iCounter := "SICK_Lector_DB_5".Data.ReadingResult.iCounter, iLength := "SICK_Lector_DB_5".Data.ReadingResult.iLength, Error_Code := "SICK_Lector_DB_5".Errorcode, Test_Comm_HMI := "BCD_Test_Comm_HMI(5)", Enable_HMI := "BCD_Enable_Trigger_HMI(5)", Disable_HMI := "BCD_Disable_Trigger_HMI(5)", Auto_Start_Lector := "Auto_Start_Lector(5)", Auto_Stop_Lector := "Auto_Stop_Lector(5)", Test_Comm => "SICK_Lector_DB_5".ComTest, Enable_Trigger => "SICK_Lector_DB_5".TriggerOn, Disable_Trigger => "SICK_Lector_DB_5".TriggerOff, Enable_Req => "SICK_Lector_DB_5".Req, Result => "SICK_Lector_DB_5".Barcode_Result, Test_OK => "SICK_Lector_DB_5".Test_OK)
   END_RUNG
   // the same network as SCL:
   "SICK_Lector_FB_DB_5"(HWInputIdent := "bcodereader_5~_32_Byte_Input_(HS)_1",   // "SICK_Lector_CLV6xx_PNDP"
                         HWInputLength := "SICK_Lector_DB_5".HWInputLength,
                         HWOutputIdent := "bcodereader_5~_32_Byte_Output_(HS)_1",
                         HWOutputLength := "SICK_Lector_DB_5".HWOutputLength,
                         CANId := "SICK_Lector_DB_5".CANId,
                         TOut := "SICK_Lector_DB_5".TOut,
                         Req := "SICK_Lector_DB_5".Req,
                         TriggerOn := "SICK_Lector_DB_5".TriggerOn,
                         TriggerOff := "SICK_Lector_DB_5".TriggerOff,
                         Matchcode := "SICK_Lector_DB_5".Matchcode,
                         SavePermanent := "SICK_Lector_DB_5".SavePermanent,
                         ComTest := "SICK_Lector_DB_5".ComTest,
                         FreeCommand := "SICK_Lector_DB_5".FreeCommand,
                         Data := "SICK_Lector_DB_5".Data,
                         RdDone => "SICK_Lector_DB_5".RdDone,
                         ReqDone => "SICK_Lector_DB_5".ReqDone,
                         ReqBusy => "SICK_Lector_DB_5".ReqBusy,
                         Error => "SICK_Lector_DB_5".Error,
                         Errorcode => "SICK_Lector_DB_5".Errorcode,
                         ENO => #_w1);
   IF #_w1 THEN
       "SICK_Lector_Control_DB_5"(Rd_Done := "SICK_Lector_DB_5".RdDone,   // "SICK_Lector_Control_FB"
                               Req_Done := "SICK_Lector_DB_5".ReqDone,
                               Req_Busy := "SICK_Lector_DB_5".ReqBusy,
                               Error := "SICK_Lector_DB_5".Error,
                               arrResult := "SICK_Lector_DB_5".Data.ReadingResult.arrResult,
                               iCounter := "SICK_Lector_DB_5".Data.ReadingResult.iCounter,
                               iLength := "SICK_Lector_DB_5".Data.ReadingResult.iLength,
                               Error_Code := "SICK_Lector_DB_5".Errorcode,
                               Test_Comm_HMI := "BCD_Test_Comm_HMI(5)",
                               Enable_HMI := "BCD_Enable_Trigger_HMI(5)",
                               Disable_HMI := "BCD_Disable_Trigger_HMI(5)",
                               Auto_Start_Lector := "Auto_Start_Lector(5)",
                               Auto_Stop_Lector := "Auto_Stop_Lector(5)",
                               Test_Comm => "SICK_Lector_DB_5".ComTest,
                               Enable_Trigger => "SICK_Lector_DB_5".TriggerOn,
                               Disable_Trigger => "SICK_Lector_DB_5".TriggerOff,
                               Enable_Req => "SICK_Lector_DB_5".Req,
                               Result => "SICK_Lector_DB_5".Barcode_Result,
                               Test_OK => "SICK_Lector_DB_5".Test_OK);
   END_IF;
END_REGION

REGION Network 46: Barcode Stations
   RUNG wire#powerrail
      "Barcode_FB_DB_1"(Sick_Result := "SICK_Lector_DB_1".Barcode_Result, Station_Control := "Control_DB".VTDBarcode_Station[1], Auto_Start_Lector := "Auto_Start_Lector(1)", Auto_Stop_Lector := "Auto_Stop_Lector(1)", "Counter" =>)
      "Barcode_FB_DB_2"(Sick_Result := "SICK_Lector_DB_2".Barcode_Result, Station_Control := "Control_DB".VTDBarcode_Station[2], Auto_Start_Lector := "Auto_Start_Lector(2)", Auto_Stop_Lector := "Auto_Stop_Lector(2)", "Counter" =>)
   END_RUNG
   RUNG wire#powerrail
      "Barcode_FB_DB_3"(Sick_Result := "SICK_Lector_DB_3".Barcode_Result, Station_Control := "Control_DB".VTDBarcode_Station[3], Auto_Start_Lector := "Auto_Start_Lector(3)", Auto_Stop_Lector := "Auto_Stop_Lector(3)", "Counter" =>)
      "Barcode_FB_DB_4"(Sick_Result := "SICK_Lector_DB_4".Barcode_Result, Station_Control := "Control_DB".VTDBarcode_Station[4], Auto_Start_Lector := "Auto_Start_Lector(4)", Auto_Stop_Lector := "Auto_Stop_Lector(4)", "Counter" =>)
   END_RUNG
   RUNG wire#powerrail
      "Barcode_FB_DB_5"(Sick_Result := "SICK_Lector_DB_5".Barcode_Result, Station_Control := "Control_DB".VTDBarcode_Station[5], Auto_Start_Lector := "Auto_Start_Lector(5)", Auto_Stop_Lector := "Auto_Stop_Lector(5)", "Counter" =>)
   END_RUNG
   // the same network as SCL:
   "Barcode_FB_DB_1"(Sick_Result := "SICK_Lector_DB_1".Barcode_Result,   // "Barcode_Station_FB"
                     Station_Control := "Control_DB".VTDBarcode_Station[1],
                     Auto_Start_Lector := "Auto_Start_Lector(1)",
                     Auto_Stop_Lector := "Auto_Stop_Lector(1)",
                     ENO => #_w1);
   IF #_w1 THEN
       "Barcode_FB_DB_2"(Sick_Result := "SICK_Lector_DB_2".Barcode_Result,   // "Barcode_Station_FB"
                         Station_Control := "Control_DB".VTDBarcode_Station[2],
                         Auto_Start_Lector := "Auto_Start_Lector(2)",
                         Auto_Stop_Lector := "Auto_Stop_Lector(2)");
   END_IF;
   "Barcode_FB_DB_3"(Sick_Result := "SICK_Lector_DB_3".Barcode_Result,   // "Barcode_Station_FB"
                     Station_Control := "Control_DB".VTDBarcode_Station[3],
                     Auto_Start_Lector := "Auto_Start_Lector(3)",
                     Auto_Stop_Lector := "Auto_Stop_Lector(3)",
                     ENO => #_w2);
   IF #_w2 THEN
       "Barcode_FB_DB_4"(Sick_Result := "SICK_Lector_DB_4".Barcode_Result,   // "Barcode_Station_FB"
                         Station_Control := "Control_DB".VTDBarcode_Station[4],
                         Auto_Start_Lector := "Auto_Start_Lector(4)",
                         Auto_Stop_Lector := "Auto_Stop_Lector(4)");
   END_IF;
   "Barcode_FB_DB_5"(Sick_Result := "SICK_Lector_DB_5".Barcode_Result,   // "Barcode_Station_FB"
                     Station_Control := "Control_DB".VTDBarcode_Station[5],
                     Auto_Start_Lector := "Auto_Start_Lector(5)",
                     Auto_Stop_Lector := "Auto_Stop_Lector(5)");
END_REGION

REGION Network 47: Stack Lights
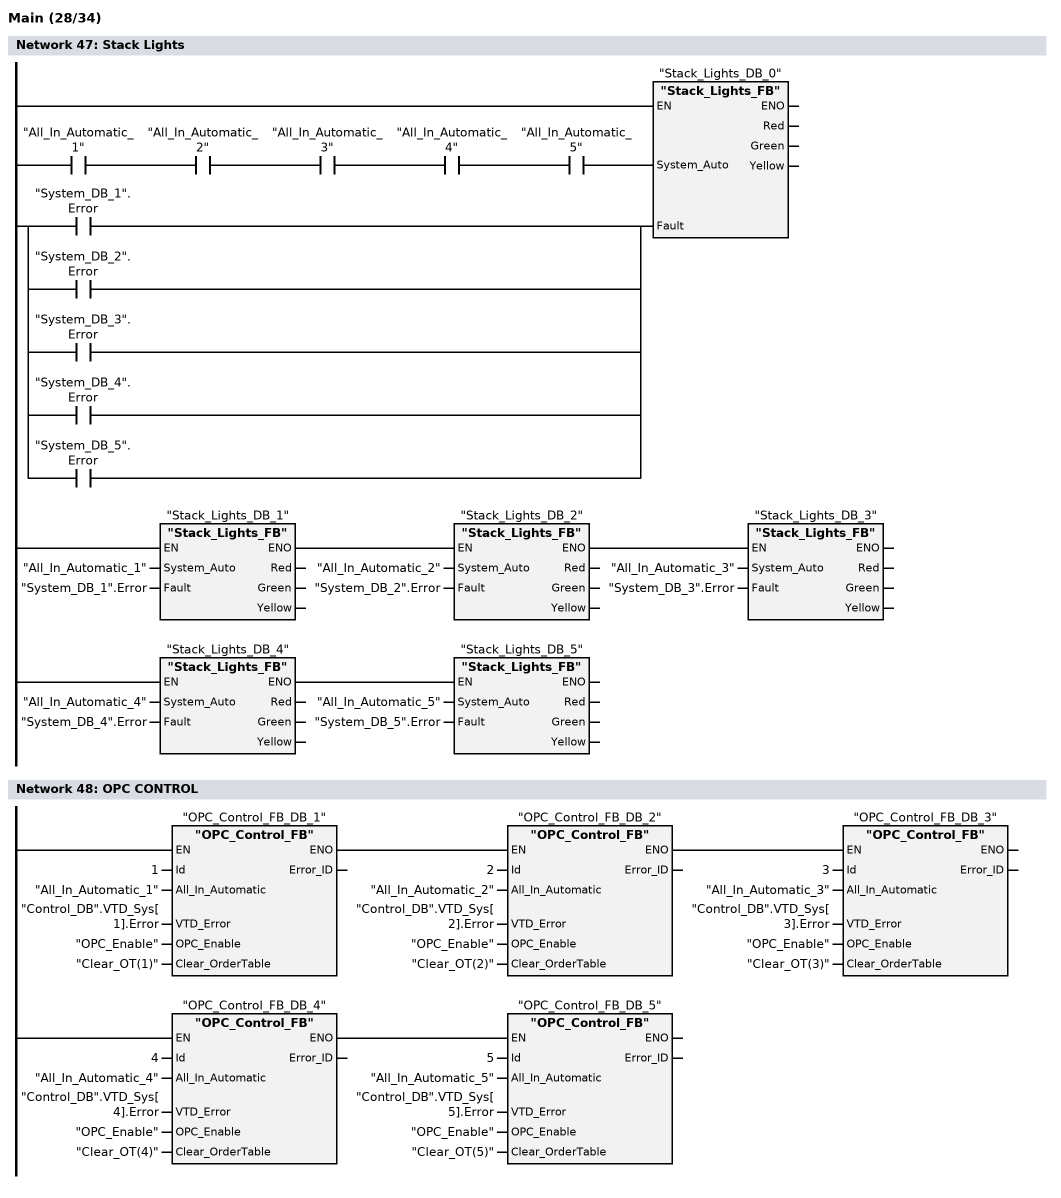
   RUNG wire#powerrail
      "Stack_Lights_DB_0"(System_Auto := wire#w1, Fault := wire#w2, Red =>, Green =>, Yellow =>)
   END_RUNG
   RUNG wire#powerrail
      Contact( "All_In_Automatic_1" )
      Contact( "All_In_Automatic_2" )
      Contact( "All_In_Automatic_3" )
      Contact( "All_In_Automatic_4" )
      Contact( "All_In_Automatic_5" )
   END_RUNG wire#w1
   RUNG wire#powerrail
      Contact( "System_DB_1".Error )
   END_RUNG wire#w2
   RUNG wire#powerrail
      Contact( "System_DB_2".Error )
   END_RUNG wire#w2
   RUNG wire#powerrail
      Contact( "System_DB_3".Error )
   END_RUNG wire#w2
   RUNG wire#powerrail
      Contact( "System_DB_4".Error )
   END_RUNG wire#w2
   RUNG wire#powerrail
      Contact( "System_DB_5".Error )
   END_RUNG wire#w2
   RUNG wire#powerrail
      "Stack_Lights_DB_1"(System_Auto := "All_In_Automatic_1", Fault := "System_DB_1".Error, Red =>, Green =>, Yellow =>)
      "Stack_Lights_DB_2"(System_Auto := "All_In_Automatic_2", Fault := "System_DB_2".Error, Red =>, Green =>, Yellow =>)
      "Stack_Lights_DB_3"(System_Auto := "All_In_Automatic_3", Fault := "System_DB_3".Error, Red =>, Green =>, Yellow =>)
   END_RUNG
   RUNG wire#powerrail
      "Stack_Lights_DB_4"(System_Auto := "All_In_Automatic_4", Fault := "System_DB_4".Error, Red =>, Green =>, Yellow =>)
      "Stack_Lights_DB_5"(System_Auto := "All_In_Automatic_5", Fault := "System_DB_5".Error, Red =>, Green =>, Yellow =>)
   END_RUNG
   // the same network as SCL:
   "Stack_Lights_DB_0"(System_Auto := "All_In_Automatic_1" AND "All_In_Automatic_2" AND "All_In_Automatic_3" AND "All_In_Automatic_4" AND "All_In_Automatic_5",   // "Stack_Lights_FB"
                       Fault := "System_DB_1".Error OR "System_DB_2".Error OR "System_DB_3".Error OR "System_DB_4".Error OR "System_DB_5".Error);
   "Stack_Lights_DB_1"(System_Auto := "All_In_Automatic_1", Fault := "System_DB_1".Error, ENO => #_w1);   // "Stack_Lights_FB"
   "Stack_Lights_DB_2"(EN := #_w1,   // "Stack_Lights_FB"
                       System_Auto := "All_In_Automatic_2",
                       Fault := "System_DB_2".Error,
                       ENO => #_w2);
   IF #_w2 THEN
       "Stack_Lights_DB_3"(System_Auto := "All_In_Automatic_3", Fault := "System_DB_3".Error);   // "Stack_Lights_FB"
   END_IF;
   "Stack_Lights_DB_4"(System_Auto := "All_In_Automatic_4", Fault := "System_DB_4".Error, ENO => #_w3);   // "Stack_Lights_FB"
   IF #_w3 THEN
       "Stack_Lights_DB_5"(System_Auto := "All_In_Automatic_5", Fault := "System_DB_5".Error);   // "Stack_Lights_FB"
   END_IF;
END_REGION

REGION Network 48: OPC CONTROL
   RUNG wire#powerrail
      "OPC_Control_FB_DB_1"(Id := 1, All_In_Automatic := "All_In_Automatic_1", VTD_Error := "Control_DB".VTD_Sys[1].Error, OPC_Enable := "OPC_Enable", Clear_OrderTable := "Clear_OT(1)", Error_ID =>)
      "OPC_Control_FB_DB_2"(Id := 2, All_In_Automatic := "All_In_Automatic_2", VTD_Error := "Control_DB".VTD_Sys[2].Error, OPC_Enable := "OPC_Enable", Clear_OrderTable := "Clear_OT(2)", Error_ID =>)
      "OPC_Control_FB_DB_3"(Id := 3, All_In_Automatic := "All_In_Automatic_3", VTD_Error := "Control_DB".VTD_Sys[3].Error, OPC_Enable := "OPC_Enable", Clear_OrderTable := "Clear_OT(3)", Error_ID =>)
   END_RUNG
   RUNG wire#powerrail
      "OPC_Control_FB_DB_4"(Id := 4, All_In_Automatic := "All_In_Automatic_4", VTD_Error := "Control_DB".VTD_Sys[4].Error, OPC_Enable := "OPC_Enable", Clear_OrderTable := "Clear_OT(4)", Error_ID =>)
      "OPC_Control_FB_DB_5"(Id := 5, All_In_Automatic := "All_In_Automatic_5", VTD_Error := "Control_DB".VTD_Sys[5].Error, OPC_Enable := "OPC_Enable", Clear_OrderTable := "Clear_OT(5)", Error_ID =>)
   END_RUNG
   // the same network as SCL:
   "OPC_Control_FB_DB_1"(Id := 1,   // "OPC_Control_FB"
                         All_In_Automatic := "All_In_Automatic_1",
                         VTD_Error := "Control_DB".VTD_Sys[1].Error,
                         OPC_Enable := "OPC_Enable",
                         Clear_OrderTable := "Clear_OT(1)",
                         ENO => #_w1);
   "OPC_Control_FB_DB_2"(EN := #_w1,   // "OPC_Control_FB"
                         Id := 2,
                         All_In_Automatic := "All_In_Automatic_2",
                         VTD_Error := "Control_DB".VTD_Sys[2].Error,
                         OPC_Enable := "OPC_Enable",
                         Clear_OrderTable := "Clear_OT(2)",
                         ENO => #_w2);
   IF #_w2 THEN
       "OPC_Control_FB_DB_3"(Id := 3,   // "OPC_Control_FB"
                             All_In_Automatic := "All_In_Automatic_3",
                             VTD_Error := "Control_DB".VTD_Sys[3].Error,
                             OPC_Enable := "OPC_Enable",
                             Clear_OrderTable := "Clear_OT(3)");
   END_IF;
   "OPC_Control_FB_DB_4"(Id := 4,   // "OPC_Control_FB"
                         All_In_Automatic := "All_In_Automatic_4",
                         VTD_Error := "Control_DB".VTD_Sys[4].Error,
                         OPC_Enable := "OPC_Enable",
                         Clear_OrderTable := "Clear_OT(4)",
                         ENO => #_w3);
   IF #_w3 THEN
       "OPC_Control_FB_DB_5"(Id := 5,   // "OPC_Control_FB"
                             All_In_Automatic := "All_In_Automatic_5",
                             VTD_Error := "Control_DB".VTD_Sys[5].Error,
                             OPC_Enable := "OPC_Enable",
                             Clear_OrderTable := "Clear_OT(5)");
   END_IF;
END_REGION

